// --- Siemens Structured Format ---
DATA_BLOCK "model_HS16_IW10"
{ S7_Optimized_Access := 'TRUE' }
VERSION : 0.1
NON_RETAIN
   VAR
      W_i : ARRAY[0..15, 0..39] OF REAL;
      W_f : ARRAY[0..15, 0..39] OF REAL;
      W_g : ARRAY[0..15, 0..39] OF REAL;
      W_o : ARRAY[0..15, 0..39] OF REAL;
      R_i : ARRAY[0..15, 0..15] OF REAL;
      R_f : ARRAY[0..15, 0..15] OF REAL;
      R_g : ARRAY[0..15, 0..15] OF REAL;
      R_o : ARRAY[0..15, 0..15] OF REAL;
      B_i : ARRAY[0..15] OF REAL;
      B_f : ARRAY[0..15] OF REAL;
      B_g : ARRAY[0..15] OF REAL;
      B_o : ARRAY[0..15] OF REAL;
      FC_W : ARRAY[0..39, 0..15] OF REAL;
      FC_B : ARRAY[0..39] OF REAL;
   END_VAR
BEGIN

      W_i[0,0] := 0.03254747;
      W_i[0,1] := 0.12385904;
      W_i[0,2] := 0.04015401;
      W_i[0,3] := -0.03803189;
      W_i[0,4] := 0.17593189;
      W_i[0,5] := 0.00417833;
      W_i[0,6] := -0.00157293;
      W_i[0,7] := 0.07286220;
      W_i[0,8] := 0.06175515;
      W_i[0,9] := -0.03080547;
      W_i[0,10] := 0.01361996;
      W_i[0,11] := -0.23670040;
      W_i[0,12] := 0.12512483;
      W_i[0,13] := -0.12038948;
      W_i[0,14] := 0.05234820;
      W_i[0,15] := 0.26305324;
      W_i[0,16] := -0.11475044;
      W_i[0,17] := 0.05957858;
      W_i[0,18] := -0.02271187;
      W_i[0,19] := -0.04982074;
      W_i[0,20] := 0.01270425;
      W_i[0,21] := 0.36205307;
      W_i[0,22] := -0.29144672;
      W_i[0,23] := 0.02366253;
      W_i[0,24] := -0.60242903;
      W_i[0,25] := -0.51985335;
      W_i[0,26] := 0.01890776;
      W_i[0,27] := -0.42442557;
      W_i[0,28] := 0.09802054;
      W_i[0,29] := -0.29197305;
      W_i[0,30] := 0.17564484;
      W_i[0,31] := -0.06584074;
      W_i[0,32] := 0.04272554;
      W_i[0,33] := 0.06813997;
      W_i[0,34] := 0.12439077;
      W_i[0,35] := -0.20625667;
      W_i[0,36] := 0.05875245;
      W_i[0,37] := -0.27000934;
      W_i[0,38] := 0.22123174;
      W_i[0,39] := 1.45426822;
      W_i[1,0] := 0.04402059;
      W_i[1,1] := 0.10076170;
      W_i[1,2] := -0.00997876;
      W_i[1,3] := 0.00796912;
      W_i[1,4] := -0.00383734;
      W_i[1,5] := -0.00800767;
      W_i[1,6] := 0.12291239;
      W_i[1,7] := 0.04417216;
      W_i[1,8] := -0.00160155;
      W_i[1,9] := -0.03973384;
      W_i[1,10] := -0.05576275;
      W_i[1,11] := 0.01415846;
      W_i[1,12] := -0.11022115;
      W_i[1,13] := 0.03613710;
      W_i[1,14] := -0.00464776;
      W_i[1,15] := -0.02071899;
      W_i[1,16] := 0.01651780;
      W_i[1,17] := -0.00011115;
      W_i[1,18] := 0.04986879;
      W_i[1,19] := -0.05042609;
      W_i[1,20] := 0.08610544;
      W_i[1,21] := 0.05673008;
      W_i[1,22] := -0.00434864;
      W_i[1,23] := 0.01197722;
      W_i[1,24] := -0.54585391;
      W_i[1,25] := -0.68996310;
      W_i[1,26] := 0.01104975;
      W_i[1,27] := 0.01825110;
      W_i[1,28] := 0.04478757;
      W_i[1,29] := -0.05586376;
      W_i[1,30] := 0.02979602;
      W_i[1,31] := 0.00707946;
      W_i[1,32] := 0.14649346;
      W_i[1,33] := 0.04832766;
      W_i[1,34] := -0.92027420;
      W_i[1,35] := -0.19189121;
      W_i[1,36] := 0.02485085;
      W_i[1,37] := -0.05241579;
      W_i[1,38] := 0.01553158;
      W_i[1,39] := -0.00394726;
      W_i[2,0] := 0.06704360;
      W_i[2,1] := -0.11752029;
      W_i[2,2] := 0.02326228;
      W_i[2,3] := -0.14317727;
      W_i[2,4] := -0.05582308;
      W_i[2,5] := 0.03605313;
      W_i[2,6] := 0.04952687;
      W_i[2,7] := -0.05419854;
      W_i[2,8] := -0.00077774;
      W_i[2,9] := 0.17699891;
      W_i[2,10] := 0.02469403;
      W_i[2,11] := 0.28494063;
      W_i[2,12] := -0.27127108;
      W_i[2,13] := -0.06837726;
      W_i[2,14] := 0.00509281;
      W_i[2,15] := 0.07467768;
      W_i[2,16] := 0.01470727;
      W_i[2,17] := 0.11394187;
      W_i[2,18] := -0.03895494;
      W_i[2,19] := 0.02999579;
      W_i[2,20] := 0.01967140;
      W_i[2,21] := 0.00220801;
      W_i[2,22] := -0.33803001;
      W_i[2,23] := 0.09799825;
      W_i[2,24] := -0.59557176;
      W_i[2,25] := -0.72284853;
      W_i[2,26] := 0.07928592;
      W_i[2,27] := -0.03053538;
      W_i[2,28] := -0.13099378;
      W_i[2,29] := -0.04490006;
      W_i[2,30] := 0.05262627;
      W_i[2,31] := -0.03356259;
      W_i[2,32] := 0.06378829;
      W_i[2,33] := -0.00362085;
      W_i[2,34] := -0.65794659;
      W_i[2,35] := 0.02030313;
      W_i[2,36] := 0.05807094;
      W_i[2,37] := -0.11176150;
      W_i[2,38] := 0.09806133;
      W_i[2,39] := -0.04513157;
      W_i[3,0] := -0.03288125;
      W_i[3,1] := 0.03644303;
      W_i[3,2] := -0.02111984;
      W_i[3,3] := -0.09554495;
      W_i[3,4] := 0.47103399;
      W_i[3,5] := -0.01821760;
      W_i[3,6] := -0.01296977;
      W_i[3,7] := 0.09772011;
      W_i[3,8] := 0.02375359;
      W_i[3,9] := 0.08029480;
      W_i[3,10] := 0.06341432;
      W_i[3,11] := -0.05777879;
      W_i[3,12] := 0.09200994;
      W_i[3,13] := -0.00543420;
      W_i[3,14] := -0.11079636;
      W_i[3,15] := 0.18567836;
      W_i[3,16] := -0.01795590;
      W_i[3,17] := -0.01424691;
      W_i[3,18] := 0.02418556;
      W_i[3,19] := -0.08783326;
      W_i[3,20] := 0.05560731;
      W_i[3,21] := 0.29868218;
      W_i[3,22] := -0.22202586;
      W_i[3,23] := -0.03734203;
      W_i[3,24] := 0.08825689;
      W_i[3,25] := 0.18388928;
      W_i[3,26] := 0.11525851;
      W_i[3,27] := -0.44497600;
      W_i[3,28] := 0.10198013;
      W_i[3,29] := -0.44026142;
      W_i[3,30] := -0.20704049;
      W_i[3,31] := 0.00454621;
      W_i[3,32] := -0.03864358;
      W_i[3,33] := -0.10321955;
      W_i[3,34] := 0.61782306;
      W_i[3,35] := -0.01621445;
      W_i[3,36] := 0.06078746;
      W_i[3,37] := 0.07829241;
      W_i[3,38] := 0.08872399;
      W_i[3,39] := 0.01815886;
      W_i[4,0] := -0.09336383;
      W_i[4,1] := 0.00870158;
      W_i[4,2] := -0.05045110;
      W_i[4,3] := 0.06854370;
      W_i[4,4] := 0.06657482;
      W_i[4,5] := -0.04358229;
      W_i[4,6] := 0.01173393;
      W_i[4,7] := 0.02832152;
      W_i[4,8] := -0.23808675;
      W_i[4,9] := 0.25903443;
      W_i[4,10] := -0.02959821;
      W_i[4,11] := -0.19702840;
      W_i[4,12] := -0.04782372;
      W_i[4,13] := 0.00693473;
      W_i[4,14] := 0.00193878;
      W_i[4,15] := 0.03396931;
      W_i[4,16] := -0.03933699;
      W_i[4,17] := -0.09345319;
      W_i[4,18] := 0.85718733;
      W_i[4,19] := -0.20839401;
      W_i[4,20] := -0.00447866;
      W_i[4,21] := -0.04350503;
      W_i[4,22] := 0.09176219;
      W_i[4,23] := 0.04992297;
      W_i[4,24] := -0.45042995;
      W_i[4,25] := 0.01641427;
      W_i[4,26] := -0.18378316;
      W_i[4,27] := 0.03955682;
      W_i[4,28] := -0.06913128;
      W_i[4,29] := 0.08025265;
      W_i[4,30] := -0.11622916;
      W_i[4,31] := 0.04558431;
      W_i[4,32] := 0.07176397;
      W_i[4,33] := -0.04032118;
      W_i[4,34] := 0.20981206;
      W_i[4,35] := -0.11253353;
      W_i[4,36] := -0.01868857;
      W_i[4,37] := -0.07242457;
      W_i[4,38] := -0.13242386;
      W_i[4,39] := -0.04244877;
      W_i[5,0] := 0.01391891;
      W_i[5,1] := -0.11018298;
      W_i[5,2] := -0.00893384;
      W_i[5,3] := -0.01407803;
      W_i[5,4] := 0.08575681;
      W_i[5,5] := 0.08241521;
      W_i[5,6] := -0.06153676;
      W_i[5,7] := 0.03060099;
      W_i[5,8] := -0.03490681;
      W_i[5,9] := 0.03142790;
      W_i[5,10] := -0.02459875;
      W_i[5,11] := 0.10959067;
      W_i[5,12] := -0.02965787;
      W_i[5,13] := 0.00184801;
      W_i[5,14] := 0.02055808;
      W_i[5,15] := -0.00937524;
      W_i[5,16] := -0.01257727;
      W_i[5,17] := 0.01791891;
      W_i[5,18] := -0.01156250;
      W_i[5,19] := -0.02731706;
      W_i[5,20] := 0.08900256;
      W_i[5,21] := 0.09895428;
      W_i[5,22] := 0.02720478;
      W_i[5,23] := 0.04369688;
      W_i[5,24] := -1.90607393;
      W_i[5,25] := -0.09418426;
      W_i[5,26] := -0.01059700;
      W_i[5,27] := -0.09780212;
      W_i[5,28] := 0.11255830;
      W_i[5,29] := 0.08197493;
      W_i[5,30] := -0.08072126;
      W_i[5,31] := 0.03083795;
      W_i[5,32] := 0.06895962;
      W_i[5,33] := 0.00149198;
      W_i[5,34] := 0.30098182;
      W_i[5,35] := 0.14424579;
      W_i[5,36] := -0.02817895;
      W_i[5,37] := -0.08498497;
      W_i[5,38] := 0.03758771;
      W_i[5,39] := 0.01095005;
      W_i[6,0] := 0.08324189;
      W_i[6,1] := -0.28836685;
      W_i[6,2] := -0.00092833;
      W_i[6,3] := -0.00874277;
      W_i[6,4] := 0.11969821;
      W_i[6,5] := -0.11207853;
      W_i[6,6] := -0.00877090;
      W_i[6,7] := -0.03745995;
      W_i[6,8] := 0.00287988;
      W_i[6,9] := 0.00178848;
      W_i[6,10] := 0.03823818;
      W_i[6,11] := 0.02621512;
      W_i[6,12] := -0.28842098;
      W_i[6,13] := -0.07084718;
      W_i[6,14] := 0.04070705;
      W_i[6,15] := -0.02042400;
      W_i[6,16] := -0.00164282;
      W_i[6,17] := 0.01065832;
      W_i[6,18] := 0.00655926;
      W_i[6,19] := 0.02358968;
      W_i[6,20] := 0.13037887;
      W_i[6,21] := 0.03868100;
      W_i[6,22] := -0.06235948;
      W_i[6,23] := 0.07983913;
      W_i[6,24] := -0.24280079;
      W_i[6,25] := -0.05732525;
      W_i[6,26] := 0.16517149;
      W_i[6,27] := -0.07414961;
      W_i[6,28] := 0.06032364;
      W_i[6,29] := 0.08282514;
      W_i[6,30] := -0.01358633;
      W_i[6,31] := 0.04311090;
      W_i[6,32] := 0.03472897;
      W_i[6,33] := -0.04253995;
      W_i[6,34] := 0.01447233;
      W_i[6,35] := 0.03594886;
      W_i[6,36] := -0.01385077;
      W_i[6,37] := 0.11164505;
      W_i[6,38] := 0.12532353;
      W_i[6,39] := -0.03726343;
      W_i[7,0] := 0.01927893;
      W_i[7,1] := 0.05625859;
      W_i[7,2] := 0.04672581;
      W_i[7,3] := -0.00316564;
      W_i[7,4] := 0.09401099;
      W_i[7,5] := -0.02755413;
      W_i[7,6] := -0.03952036;
      W_i[7,7] := 0.03364034;
      W_i[7,8] := 0.05500693;
      W_i[7,9] := 0.02471298;
      W_i[7,10] := 0.03820876;
      W_i[7,11] := -0.26921606;
      W_i[7,12] := -0.02231521;
      W_i[7,13] := -0.01752430;
      W_i[7,14] := 0.03934914;
      W_i[7,15] := 0.01282423;
      W_i[7,16] := -0.08716010;
      W_i[7,17] := -0.09125534;
      W_i[7,18] := 0.00613662;
      W_i[7,19] := 0.08651425;
      W_i[7,20] := -0.01288831;
      W_i[7,21] := 0.20176773;
      W_i[7,22] := -0.20166723;
      W_i[7,23] := 0.01241351;
      W_i[7,24] := -0.87556225;
      W_i[7,25] := -0.46218389;
      W_i[7,26] := 0.09773878;
      W_i[7,27] := -0.12810560;
      W_i[7,28] := 0.04194518;
      W_i[7,29] := -0.03563948;
      W_i[7,30] := 0.08049577;
      W_i[7,31] := 0.04509509;
      W_i[7,32] := -0.11332804;
      W_i[7,33] := 0.10539962;
      W_i[7,34] := 0.24167158;
      W_i[7,35] := 0.04508473;
      W_i[7,36] := 0.00324964;
      W_i[7,37] := 0.22550038;
      W_i[7,38] := 0.17509922;
      W_i[7,39] := -0.77876335;
      W_i[8,0] := -0.03076644;
      W_i[8,1] := 0.03958185;
      W_i[8,2] := 0.05958826;
      W_i[8,3] := 0.00143461;
      W_i[8,4] := -0.03551066;
      W_i[8,5] := 0.06705590;
      W_i[8,6] := -0.00545013;
      W_i[8,7] := -0.11520024;
      W_i[8,8] := -0.04941865;
      W_i[8,9] := 0.00970779;
      W_i[8,10] := -0.02700928;
      W_i[8,11] := 0.12616971;
      W_i[8,12] := -0.23012702;
      W_i[8,13] := -0.13218109;
      W_i[8,14] := 0.10565390;
      W_i[8,15] := 0.03265957;
      W_i[8,16] := 0.01893855;
      W_i[8,17] := 0.05783269;
      W_i[8,18] := 0.04541522;
      W_i[8,19] := -0.17565091;
      W_i[8,20] := -0.03008310;
      W_i[8,21] := 0.02609591;
      W_i[8,22] := -0.11792074;
      W_i[8,23] := -0.03097328;
      W_i[8,24] := -1.12349439;
      W_i[8,25] := -0.10578562;
      W_i[8,26] := 0.11967086;
      W_i[8,27] := -0.19309855;
      W_i[8,28] := -0.04314341;
      W_i[8,29] := -0.02280886;
      W_i[8,30] := 0.09419166;
      W_i[8,31] := -0.00168002;
      W_i[8,32] := 0.17011297;
      W_i[8,33] := 0.12776379;
      W_i[8,34] := 0.00792190;
      W_i[8,35] := 0.00793266;
      W_i[8,36] := 0.02933485;
      W_i[8,37] := -0.04765635;
      W_i[8,38] := -0.05385318;
      W_i[8,39] := 1.04576063;
      W_i[9,0] := 0.15918908;
      W_i[9,1] := 0.04106269;
      W_i[9,2] := 0.02940365;
      W_i[9,3] := -0.02633034;
      W_i[9,4] := 0.06646424;
      W_i[9,5] := -0.06870057;
      W_i[9,6] := 0.00617184;
      W_i[9,7] := 0.01493581;
      W_i[9,8] := 0.00472299;
      W_i[9,9] := -0.18171085;
      W_i[9,10] := -0.00863580;
      W_i[9,11] := 0.11203966;
      W_i[9,12] := 0.03235663;
      W_i[9,13] := -0.00635904;
      W_i[9,14] := -0.00805719;
      W_i[9,15] := 0.03256573;
      W_i[9,16] := -0.02982800;
      W_i[9,17] := 0.02432551;
      W_i[9,18] := -0.04791717;
      W_i[9,19] := -0.03479305;
      W_i[9,20] := 0.02419964;
      W_i[9,21] := -0.00806570;
      W_i[9,22] := 0.00884045;
      W_i[9,23] := 0.00822151;
      W_i[9,24] := -0.46266055;
      W_i[9,25] := -0.24154246;
      W_i[9,26] := 0.10637723;
      W_i[9,27] := 0.00555547;
      W_i[9,28] := 0.00231378;
      W_i[9,29] := 0.17306480;
      W_i[9,30] := -0.14428723;
      W_i[9,31] := -0.01611738;
      W_i[9,32] := -0.15273547;
      W_i[9,33] := -0.03995335;
      W_i[9,34] := -0.60233766;
      W_i[9,35] := -0.06071381;
      W_i[9,36] := 0.01153921;
      W_i[9,37] := 0.15725203;
      W_i[9,38] := 0.04887648;
      W_i[9,39] := 0.03194974;
      W_i[10,0] := 0.00000571;
      W_i[10,1] := 0.02921890;
      W_i[10,2] := 0.03921259;
      W_i[10,3] := -0.10342362;
      W_i[10,4] := 0.04451175;
      W_i[10,5] := -0.01788418;
      W_i[10,6] := 0.06014212;
      W_i[10,7] := -0.12761596;
      W_i[10,8] := 0.10969678;
      W_i[10,9] := 0.13464272;
      W_i[10,10] := -0.07629871;
      W_i[10,11] := -1.31473470;
      W_i[10,12] := 0.97041023;
      W_i[10,13] := -0.02917644;
      W_i[10,14] := 0.26857987;
      W_i[10,15] := 0.06801854;
      W_i[10,16] := -0.22419471;
      W_i[10,17] := 0.26248446;
      W_i[10,18] := -0.16949444;
      W_i[10,19] := -0.11971024;
      W_i[10,20] := -0.15914336;
      W_i[10,21] := 0.18180194;
      W_i[10,22] := -0.44877753;
      W_i[10,23] := 0.05718501;
      W_i[10,24] := 0.77401525;
      W_i[10,25] := 0.61128056;
      W_i[10,26] := 0.00735129;
      W_i[10,27] := -0.08243502;
      W_i[10,28] := -0.03729297;
      W_i[10,29] := 0.16128409;
      W_i[10,30] := -0.02351914;
      W_i[10,31] := 0.10431249;
      W_i[10,32] := 0.05746254;
      W_i[10,33] := 0.08887602;
      W_i[10,34] := -0.39106452;
      W_i[10,35] := 0.22569241;
      W_i[10,36] := -0.13208193;
      W_i[10,37] := -0.16115883;
      W_i[10,38] := 0.27080455;
      W_i[10,39] := 0.62801355;
      W_i[11,0] := -0.05849513;
      W_i[11,1] := -0.03062119;
      W_i[11,2] := -0.00411083;
      W_i[11,3] := 0.00799791;
      W_i[11,4] := 0.08333463;
      W_i[11,5] := 0.02937987;
      W_i[11,6] := 0.06844535;
      W_i[11,7] := -0.01198280;
      W_i[11,8] := 0.05660131;
      W_i[11,9] := -0.14609326;
      W_i[11,10] := -0.01666861;
      W_i[11,11] := -0.06908122;
      W_i[11,12] := 0.15483312;
      W_i[11,13] := -0.00687739;
      W_i[11,14] := 0.01971146;
      W_i[11,15] := 0.13305922;
      W_i[11,16] := -0.02189317;
      W_i[11,17] := 0.00985993;
      W_i[11,18] := -0.14880668;
      W_i[11,19] := 0.01909257;
      W_i[11,20] := 0.03714932;
      W_i[11,21] := -0.02673176;
      W_i[11,22] := -0.02788893;
      W_i[11,23] := 0.11408952;
      W_i[11,24] := -0.37118840;
      W_i[11,25] := -0.08985706;
      W_i[11,26] := -0.11023268;
      W_i[11,27] := 0.05117378;
      W_i[11,28] := 0.08547711;
      W_i[11,29] := 0.12702477;
      W_i[11,30] := 0.10544877;
      W_i[11,31] := -0.00480978;
      W_i[11,32] := 0.16144946;
      W_i[11,33] := 0.05210381;
      W_i[11,34] := -0.00085451;
      W_i[11,35] := -0.00874526;
      W_i[11,36] := -0.06161120;
      W_i[11,37] := -0.36774832;
      W_i[11,38] := 0.04212995;
      W_i[11,39] := 0.03037546;
      W_i[12,0] := 0.00629061;
      W_i[12,1] := -0.06136212;
      W_i[12,2] := -0.00718669;
      W_i[12,3] := -0.10042179;
      W_i[12,4] := 0.06293897;
      W_i[12,5] := -0.03143417;
      W_i[12,6] := -0.03538829;
      W_i[12,7] := 0.07763195;
      W_i[12,8] := -0.01023159;
      W_i[12,9] := -0.11412965;
      W_i[12,10] := -0.01354402;
      W_i[12,11] := -0.02311977;
      W_i[12,12] := 0.02796080;
      W_i[12,13] := 0.07165248;
      W_i[12,14] := -0.03632027;
      W_i[12,15] := 0.03878558;
      W_i[12,16] := -0.07312500;
      W_i[12,17] := 0.01845204;
      W_i[12,18] := -0.08527449;
      W_i[12,19] := -0.00854577;
      W_i[12,20] := 0.00351815;
      W_i[12,21] := -0.16628480;
      W_i[12,22] := 0.06705266;
      W_i[12,23] := 0.14307018;
      W_i[12,24] := -0.53957397;
      W_i[12,25] := -0.87219816;
      W_i[12,26] := -0.06440469;
      W_i[12,27] := 0.07379381;
      W_i[12,28] := 0.07828815;
      W_i[12,29] := 0.38822088;
      W_i[12,30] := 0.11594980;
      W_i[12,31] := 0.05581488;
      W_i[12,32] := 0.30664018;
      W_i[12,33] := 0.12759578;
      W_i[12,34] := -0.14797799;
      W_i[12,35] := 0.14329346;
      W_i[12,36] := 0.22981535;
      W_i[12,37] := 0.00895516;
      W_i[12,38] := 0.20012984;
      W_i[12,39] := 0.09707437;
      W_i[13,0] := 0.07871004;
      W_i[13,1] := 0.06409820;
      W_i[13,2] := -0.00181766;
      W_i[13,3] := 0.05780525;
      W_i[13,4] := 0.21016718;
      W_i[13,5] := 0.05360549;
      W_i[13,6] := -0.08758270;
      W_i[13,7] := -0.33428112;
      W_i[13,8] := -0.09135646;
      W_i[13,9] := 0.11706311;
      W_i[13,10] := -0.05231260;
      W_i[13,11] := -0.03317479;
      W_i[13,12] := -0.40338296;
      W_i[13,13] := -0.00985299;
      W_i[13,14] := 0.02202887;
      W_i[13,15] := 0.13037799;
      W_i[13,16] := 0.04808246;
      W_i[13,17] := 0.04501719;
      W_i[13,18] := -0.01153503;
      W_i[13,19] := 0.03141625;
      W_i[13,20] := 0.02999944;
      W_i[13,21] := 0.01402024;
      W_i[13,22] := 0.06788336;
      W_i[13,23] := -0.09942459;
      W_i[13,24] := 0.31843993;
      W_i[13,25] := 0.10697926;
      W_i[13,26] := -0.06989229;
      W_i[13,27] := 0.10588147;
      W_i[13,28] := 0.06872193;
      W_i[13,29] := -0.15371445;
      W_i[13,30] := 0.06626805;
      W_i[13,31] := -0.05594840;
      W_i[13,32] := -0.09573574;
      W_i[13,33] := 0.05669653;
      W_i[13,34] := 0.06202357;
      W_i[13,35] := -0.13674185;
      W_i[13,36] := 0.06451428;
      W_i[13,37] := 0.12041676;
      W_i[13,38] := -0.16850901;
      W_i[13,39] := 0.97759265;
      W_i[14,0] := 0.00773311;
      W_i[14,1] := -0.06673568;
      W_i[14,2] := -0.03463669;
      W_i[14,3] := -0.07830913;
      W_i[14,4] := 0.22799005;
      W_i[14,5] := -0.23448689;
      W_i[14,6] := 0.19569355;
      W_i[14,7] := 0.13153341;
      W_i[14,8] := -0.12420856;
      W_i[14,9] := 0.28603974;
      W_i[14,10] := -0.09231006;
      W_i[14,11] := -0.25477913;
      W_i[14,12] := 0.14903630;
      W_i[14,13] := -0.29128024;
      W_i[14,14] := 0.10725706;
      W_i[14,15] := 0.13540378;
      W_i[14,16] := -0.09035023;
      W_i[14,17] := -0.01749873;
      W_i[14,18] := -0.47894967;
      W_i[14,19] := -0.06870104;
      W_i[14,20] := -0.17096391;
      W_i[14,21] := -0.05212005;
      W_i[14,22] := -0.16184741;
      W_i[14,23] := -0.21394062;
      W_i[14,24] := -0.75706887;
      W_i[14,25] := -0.70485926;
      W_i[14,26] := -0.33521020;
      W_i[14,27] := 0.03507431;
      W_i[14,28] := -0.12678961;
      W_i[14,29] := 0.16709636;
      W_i[14,30] := -0.05052740;
      W_i[14,31] := -0.11800393;
      W_i[14,32] := -0.09575160;
      W_i[14,33] := -0.01452094;
      W_i[14,34] := 0.00625472;
      W_i[14,35] := -0.12877558;
      W_i[14,36] := -0.06069501;
      W_i[14,37] := -0.22877042;
      W_i[14,38] := 0.17231728;
      W_i[14,39] := 1.04831111;
      W_i[15,0] := 0.04376059;
      W_i[15,1] := -0.02296846;
      W_i[15,2] := 0.01713722;
      W_i[15,3] := 0.17107451;
      W_i[15,4] := 0.17369278;
      W_i[15,5] := -0.01825109;
      W_i[15,6] := -0.02258963;
      W_i[15,7] := 0.02190229;
      W_i[15,8] := -0.03702974;
      W_i[15,9] := -0.03196403;
      W_i[15,10] := 0.08264420;
      W_i[15,11] := 0.05920084;
      W_i[15,12] := -0.42805931;
      W_i[15,13] := -0.17172982;
      W_i[15,14] := 0.02115602;
      W_i[15,15] := -0.00198027;
      W_i[15,16] := 0.02912534;
      W_i[15,17] := -0.07075519;
      W_i[15,18] := -0.11744455;
      W_i[15,19] := 0.30688557;
      W_i[15,20] := 0.04301663;
      W_i[15,21] := 0.21635388;
      W_i[15,22] := -0.08966552;
      W_i[15,23] := 0.07217173;
      W_i[15,24] := -0.53244919;
      W_i[15,25] := -0.17169446;
      W_i[15,26] := -0.00556448;
      W_i[15,27] := -0.16294074;
      W_i[15,28] := 0.03264420;
      W_i[15,29] := 0.01573053;
      W_i[15,30] := -0.03329111;
      W_i[15,31] := -0.01247096;
      W_i[15,32] := 0.21000683;
      W_i[15,33] := 0.15043637;
      W_i[15,34] := -0.16979790;
      W_i[15,35] := 0.00504174;
      W_i[15,36] := 0.00267995;
      W_i[15,37] := -0.06215737;
      W_i[15,38] := 0.21481486;
      W_i[15,39] := 0.07231134;
      W_f[0,0] := -0.02091779;
      W_f[0,1] := -0.01810063;
      W_f[0,2] := 0.21008702;
      W_f[0,3] := 0.09207959;
      W_f[0,4] := -0.10695104;
      W_f[0,5] := -0.03611851;
      W_f[0,6] := 0.03397696;
      W_f[0,7] := 0.16544856;
      W_f[0,8] := -0.05997881;
      W_f[0,9] := -0.00453302;
      W_f[0,10] := 0.03307042;
      W_f[0,11] := 0.14202486;
      W_f[0,12] := 0.08012222;
      W_f[0,13] := -0.01528266;
      W_f[0,14] := -0.15201145;
      W_f[0,15] := -0.15718380;
      W_f[0,16] := -0.08413183;
      W_f[0,17] := 0.20222495;
      W_f[0,18] := -0.01353853;
      W_f[0,19] := 0.02782044;
      W_f[0,20] := -0.04748038;
      W_f[0,21] := 0.18304287;
      W_f[0,22] := 0.31257400;
      W_f[0,23] := -0.06208337;
      W_f[0,24] := 1.60133708;
      W_f[0,25] := 1.51956844;
      W_f[0,26] := 0.00266673;
      W_f[0,27] := 0.12180892;
      W_f[0,28] := 0.04435247;
      W_f[0,29] := 0.03200248;
      W_f[0,30] := 0.38338348;
      W_f[0,31] := 0.04435838;
      W_f[0,32] := 0.30680922;
      W_f[0,33] := 0.13231254;
      W_f[0,34] := 1.35719514;
      W_f[0,35] := 0.36870065;
      W_f[0,36] := 0.08067872;
      W_f[0,37] := 0.21299456;
      W_f[0,38] := -0.02734181;
      W_f[0,39] := 0.07611577;
      W_f[1,0] := -0.38817102;
      W_f[1,1] := 0.02779610;
      W_f[1,2] := -0.26510856;
      W_f[1,3] := -0.07072625;
      W_f[1,4] := 0.11966246;
      W_f[1,5] := 0.12000409;
      W_f[1,6] := -0.50846916;
      W_f[1,7] := -0.13361093;
      W_f[1,8] := -0.13777961;
      W_f[1,9] := -0.08736181;
      W_f[1,10] := 0.31134772;
      W_f[1,11] := 0.08504082;
      W_f[1,12] := 0.21148330;
      W_f[1,13] := -0.13549544;
      W_f[1,14] := -0.12279948;
      W_f[1,15] := 0.05185516;
      W_f[1,16] := -0.14745373;
      W_f[1,17] := 0.05817819;
      W_f[1,18] := 1.08165765;
      W_f[1,19] := 0.18381153;
      W_f[1,20] := 0.28742057;
      W_f[1,21] := -0.27315989;
      W_f[1,22] := 0.08855448;
      W_f[1,23] := -0.09573217;
      W_f[1,24] := -0.36683315;
      W_f[1,25] := -0.69911557;
      W_f[1,26] := 0.07979747;
      W_f[1,27] := -0.17541142;
      W_f[1,28] := -0.24551585;
      W_f[1,29] := 0.14984873;
      W_f[1,30] := 0.02324941;
      W_f[1,31] := 0.07932284;
      W_f[1,32] := -0.12442444;
      W_f[1,33] := 0.02366536;
      W_f[1,34] := 0.13745289;
      W_f[1,35] := 0.46306115;
      W_f[1,36] := -0.22673251;
      W_f[1,37] := 0.07258049;
      W_f[1,38] := 0.42296681;
      W_f[1,39] := 0.14921528;
      W_f[2,0] := -0.01982149;
      W_f[2,1] := 0.03324119;
      W_f[2,2] := -0.04425151;
      W_f[2,3] := 0.08356856;
      W_f[2,4] := -0.00266197;
      W_f[2,5] := -0.01017811;
      W_f[2,6] := -0.03237398;
      W_f[2,7] := -0.00609645;
      W_f[2,8] := -0.04705935;
      W_f[2,9] := 0.03853706;
      W_f[2,10] := 0.03140420;
      W_f[2,11] := -0.12043314;
      W_f[2,12] := 0.26915759;
      W_f[2,13] := 0.04188414;
      W_f[2,14] := 0.10631428;
      W_f[2,15] := 0.05646345;
      W_f[2,16] := 0.16197611;
      W_f[2,17] := 0.21402863;
      W_f[2,18] := -0.09279267;
      W_f[2,19] := -0.00577110;
      W_f[2,20] := -0.03028176;
      W_f[2,21] := -0.05153098;
      W_f[2,22] := -0.11017115;
      W_f[2,23] := -0.01419843;
      W_f[2,24] := -0.63084757;
      W_f[2,25] := -0.41158974;
      W_f[2,26] := -0.14941035;
      W_f[2,27] := 0.04505387;
      W_f[2,28] := 0.09163468;
      W_f[2,29] := 0.20423372;
      W_f[2,30] := -0.05021087;
      W_f[2,31] := -0.05815214;
      W_f[2,32] := -0.04207016;
      W_f[2,33] := 0.21736744;
      W_f[2,34] := 0.64307344;
      W_f[2,35] := -0.19552369;
      W_f[2,36] := -0.05630085;
      W_f[2,37] := 0.00531330;
      W_f[2,38] := -0.12282822;
      W_f[2,39] := 0.54551679;
      W_f[3,0] := -0.00758014;
      W_f[3,1] := 0.00559481;
      W_f[3,2] := 0.04034248;
      W_f[3,3] := 0.02266315;
      W_f[3,4] := -0.09543922;
      W_f[3,5] := 0.03211372;
      W_f[3,6] := 0.07329436;
      W_f[3,7] := -0.04057672;
      W_f[3,8] := -0.09598581;
      W_f[3,9] := -0.00159119;
      W_f[3,10] := 0.00039486;
      W_f[3,11] := -0.00788106;
      W_f[3,12] := -0.06210583;
      W_f[3,13] := -0.01413072;
      W_f[3,14] := -0.24013861;
      W_f[3,15] := -0.07759018;
      W_f[3,16] := 0.04360460;
      W_f[3,17] := -0.20987833;
      W_f[3,18] := 0.14860362;
      W_f[3,19] := -0.02982033;
      W_f[3,20] := -0.08417022;
      W_f[3,21] := 0.08484244;
      W_f[3,22] := 0.33418563;
      W_f[3,23] := -0.01567571;
      W_f[3,24] := 1.09344435;
      W_f[3,25] := 0.97723728;
      W_f[3,26] := -0.13622019;
      W_f[3,27] := -0.09956130;
      W_f[3,28] := 0.00698416;
      W_f[3,29] := 0.00054130;
      W_f[3,30] := 0.26053473;
      W_f[3,31] := -0.09947061;
      W_f[3,32] := 0.26287073;
      W_f[3,33] := 0.00611334;
      W_f[3,34] := 1.38905013;
      W_f[3,35] := -0.14349753;
      W_f[3,36] := -0.00342261;
      W_f[3,37] := -0.06542191;
      W_f[3,38] := 0.10482345;
      W_f[3,39] := 0.11385954;
      W_f[4,0] := 0.28678942;
      W_f[4,1] := -0.14550023;
      W_f[4,2] := 0.20301139;
      W_f[4,3] := -0.15284956;
      W_f[4,4] := -0.11934043;
      W_f[4,5] := -0.06261637;
      W_f[4,6] := -0.09047025;
      W_f[4,7] := -0.02217131;
      W_f[4,8] := 0.32893139;
      W_f[4,9] := -0.50192183;
      W_f[4,10] := -0.02496753;
      W_f[4,11] := -0.02753776;
      W_f[4,12] := -0.31547716;
      W_f[4,13] := -0.04408565;
      W_f[4,14] := 0.05384916;
      W_f[4,15] := -0.32536885;
      W_f[4,16] := -0.01380023;
      W_f[4,17] := -0.12124701;
      W_f[4,18] := 0.62146658;
      W_f[4,19] := 0.01393374;
      W_f[4,20] := 0.04359875;
      W_f[4,21] := 0.16302615;
      W_f[4,22] := -0.21024738;
      W_f[4,23] := -0.12911762;
      W_f[4,24] := -0.08685920;
      W_f[4,25] := -0.03674764;
      W_f[4,26] := 0.30872664;
      W_f[4,27] := 0.03806484;
      W_f[4,28] := 0.01020021;
      W_f[4,29] := -0.15197505;
      W_f[4,30] := 0.05839425;
      W_f[4,31] := -0.01564794;
      W_f[4,32] := -0.18343291;
      W_f[4,33] := 0.02443381;
      W_f[4,34] := 0.21402271;
      W_f[4,35] := 0.19360679;
      W_f[4,36] := 0.09160208;
      W_f[4,37] := 0.06046678;
      W_f[4,38] := -0.08968955;
      W_f[4,39] := -0.03439303;
      W_f[5,0] := -0.39957133;
      W_f[5,1] := -0.46507514;
      W_f[5,2] := -0.26463589;
      W_f[5,3] := -0.08991144;
      W_f[5,4] := -0.16602752;
      W_f[5,5] := 0.36502278;
      W_f[5,6] := -0.03514609;
      W_f[5,7] := -0.06387420;
      W_f[5,8] := 0.12637840;
      W_f[5,9] := 0.19450709;
      W_f[5,10] := -0.07852599;
      W_f[5,11] := -0.24370454;
      W_f[5,12] := -0.06879438;
      W_f[5,13] := 0.26811865;
      W_f[5,14] := 0.01808503;
      W_f[5,15] := -0.10070925;
      W_f[5,16] := 0.31043285;
      W_f[5,17] := -0.03764273;
      W_f[5,18] := -0.05466426;
      W_f[5,19] := -0.10286047;
      W_f[5,20] := -0.18913145;
      W_f[5,21] := -0.06289500;
      W_f[5,22] := 0.26261428;
      W_f[5,23] := 0.11659861;
      W_f[5,24] := 2.13931274;
      W_f[5,25] := 2.36269403;
      W_f[5,26] := -0.41290748;
      W_f[5,27] := 0.08711372;
      W_f[5,28] := -0.06960621;
      W_f[5,29] := -0.10882857;
      W_f[5,30] := 0.02405319;
      W_f[5,31] := -0.02791615;
      W_f[5,32] := -0.03174478;
      W_f[5,33] := -0.22598031;
      W_f[5,34] := 0.02213258;
      W_f[5,35] := 0.06206211;
      W_f[5,36] := -0.22062500;
      W_f[5,37] := 0.20298730;
      W_f[5,38] := 0.03730853;
      W_f[5,39] := -0.16448267;
      W_f[6,0] := 0.09157378;
      W_f[6,1] := -0.10600298;
      W_f[6,2] := 0.01516851;
      W_f[6,3] := -0.09814398;
      W_f[6,4] := -0.02060772;
      W_f[6,5] := -0.11663528;
      W_f[6,6] := 0.17605469;
      W_f[6,7] := 0.14043835;
      W_f[6,8] := -0.06626645;
      W_f[6,9] := 0.03254180;
      W_f[6,10] := -0.03667779;
      W_f[6,11] := 0.03295979;
      W_f[6,12] := 0.13456115;
      W_f[6,13] := 0.17527823;
      W_f[6,14] := 0.06438499;
      W_f[6,15] := -0.12721057;
      W_f[6,16] := -0.28780875;
      W_f[6,17] := 0.11614764;
      W_f[6,18] := -0.23114346;
      W_f[6,19] := -0.07521003;
      W_f[6,20] := -0.14160164;
      W_f[6,21] := 0.12687035;
      W_f[6,22] := 0.38557813;
      W_f[6,23] := -0.12900937;
      W_f[6,24] := 1.14550745;
      W_f[6,25] := 1.20651269;
      W_f[6,26] := 0.01718643;
      W_f[6,27] := -0.20140134;
      W_f[6,28] := -0.03907681;
      W_f[6,29] := -1.03183591;
      W_f[6,30] := 0.13298695;
      W_f[6,31] := -0.05304611;
      W_f[6,32] := 0.27542382;
      W_f[6,33] := 0.48400101;
      W_f[6,34] := 0.87303483;
      W_f[6,35] := -0.27916309;
      W_f[6,36] := 0.09285419;
      W_f[6,37] := -0.00086587;
      W_f[6,38] := 0.21403548;
      W_f[6,39] := 0.01036415;
      W_f[7,0] := -0.00185265;
      W_f[7,1] := 0.07858364;
      W_f[7,2] := 0.00610039;
      W_f[7,3] := 0.06575946;
      W_f[7,4] := -0.08100830;
      W_f[7,5] := 0.00321988;
      W_f[7,6] := 0.07597861;
      W_f[7,7] := -0.12638623;
      W_f[7,8] := 0.14672390;
      W_f[7,9] := 0.04145058;
      W_f[7,10] := 0.03552409;
      W_f[7,11] := -0.42004111;
      W_f[7,12] := 0.25357988;
      W_f[7,13] := -0.08330481;
      W_f[7,14] := -0.08974353;
      W_f[7,15] := -0.10517624;
      W_f[7,16] := -0.38224444;
      W_f[7,17] := -0.45799860;
      W_f[7,18] := -0.06309059;
      W_f[7,19] := -0.30799860;
      W_f[7,20] := -0.08522949;
      W_f[7,21] := -0.06581733;
      W_f[7,22] := 0.25805131;
      W_f[7,23] := 0.02311642;
      W_f[7,24] := 0.90950686;
      W_f[7,25] := 1.18889558;
      W_f[7,26] := -0.11546607;
      W_f[7,27] := -0.10872247;
      W_f[7,28] := -0.08876549;
      W_f[7,29] := 0.00109644;
      W_f[7,30] := 0.23372188;
      W_f[7,31] := -0.13769329;
      W_f[7,32] := 0.16597158;
      W_f[7,33] := 0.04170239;
      W_f[7,34] := 1.31133747;
      W_f[7,35] := -0.11888772;
      W_f[7,36] := 0.04907094;
      W_f[7,37] := 0.14026117;
      W_f[7,38] := 0.12559824;
      W_f[7,39] := -1.27418923;
      W_f[8,0] := 0.12555996;
      W_f[8,1] := -0.10315757;
      W_f[8,2] := 0.03551091;
      W_f[8,3] := -0.03898631;
      W_f[8,4] := -0.13206761;
      W_f[8,5] := 0.07454634;
      W_f[8,6] := 0.10206546;
      W_f[8,7] := 0.01262685;
      W_f[8,8] := -0.00534601;
      W_f[8,9] := -0.00536494;
      W_f[8,10] := -0.04092396;
      W_f[8,11] := -0.38692373;
      W_f[8,12] := 0.03422466;
      W_f[8,13] := 0.02580789;
      W_f[8,14] := 0.26898870;
      W_f[8,15] := -0.24944888;
      W_f[8,16] := -0.02722716;
      W_f[8,17] := -0.10108043;
      W_f[8,18] := 0.54244351;
      W_f[8,19] := -0.23120664;
      W_f[8,20] := -0.04103015;
      W_f[8,21] := -0.16740812;
      W_f[8,22] := 0.13893805;
      W_f[8,23] := -0.04656294;
      W_f[8,24] := 0.53174204;
      W_f[8,25] := 0.74309415;
      W_f[8,26] := -0.00084738;
      W_f[8,27] := -0.04600925;
      W_f[8,28] := -0.15880004;
      W_f[8,29] := 0.08535929;
      W_f[8,30] := 0.10221286;
      W_f[8,31] := -0.03335671;
      W_f[8,32] := 0.03138823;
      W_f[8,33] := -0.02403146;
      W_f[8,34] := 0.83305961;
      W_f[8,35] := -0.07033388;
      W_f[8,36] := -0.17499864;
      W_f[8,37] := 0.09229370;
      W_f[8,38] := -0.17668678;
      W_f[8,39] := 0.14198503;
      W_f[9,0] := -0.08198071;
      W_f[9,1] := 0.03835172;
      W_f[9,2] := 1.02026522;
      W_f[9,3] := -0.15293953;
      W_f[9,4] := -0.16179894;
      W_f[9,5] := 0.03072036;
      W_f[9,6] := -0.09759208;
      W_f[9,7] := -0.07946933;
      W_f[9,8] := -0.65491873;
      W_f[9,9] := 0.24554865;
      W_f[9,10] := -0.00084776;
      W_f[9,11] := -0.02393647;
      W_f[9,12] := -0.11035760;
      W_f[9,13] := 0.05757844;
      W_f[9,14] := 0.00252463;
      W_f[9,15] := -0.04278835;
      W_f[9,16] := -0.01363701;
      W_f[9,17] := 0.03181182;
      W_f[9,18] := 0.29542166;
      W_f[9,19] := 0.18680713;
      W_f[9,20] := -0.14596237;
      W_f[9,21] := 0.04626612;
      W_f[9,22] := -0.49596560;
      W_f[9,23] := -0.29882804;
      W_f[9,24] := -0.05025842;
      W_f[9,25] := -0.24922217;
      W_f[9,26] := 0.22770426;
      W_f[9,27] := -0.07712200;
      W_f[9,28] := -0.16018625;
      W_f[9,29] := -0.36028501;
      W_f[9,30] := -0.15894593;
      W_f[9,31] := 0.07634185;
      W_f[9,32] := -0.14248089;
      W_f[9,33] := 0.47243714;
      W_f[9,34] := 0.37227076;
      W_f[9,35] := 0.08862774;
      W_f[9,36] := 0.18020450;
      W_f[9,37] := -0.46372715;
      W_f[9,38] := 0.10143350;
      W_f[9,39] := 0.03257460;
      W_f[10,0] := 0.01476683;
      W_f[10,1] := 0.08915940;
      W_f[10,2] := 0.09493639;
      W_f[10,3] := 0.00921640;
      W_f[10,4] := -0.40101719;
      W_f[10,5] := -0.09464957;
      W_f[10,6] := -0.04691195;
      W_f[10,7] := -0.02866868;
      W_f[10,8] := -0.04315028;
      W_f[10,9] := -0.17093825;
      W_f[10,10] := -0.00073274;
      W_f[10,11] := -0.27505547;
      W_f[10,12] := 0.33605671;
      W_f[10,13] := -0.22034417;
      W_f[10,14] := 0.24165145;
      W_f[10,15] := -0.23521844;
      W_f[10,16] := -0.00154005;
      W_f[10,17] := -0.00158511;
      W_f[10,18] := 0.11912328;
      W_f[10,19] := -0.02448388;
      W_f[10,20] := -0.23859039;
      W_f[10,21] := -0.05945824;
      W_f[10,22] := 0.01714438;
      W_f[10,23] := -0.18285508;
      W_f[10,24] := 1.57859039;
      W_f[10,25] := 1.89422643;
      W_f[10,26] := 0.09559432;
      W_f[10,27] := -0.27382705;
      W_f[10,28] := -0.28146487;
      W_f[10,29] := 0.04344108;
      W_f[10,30] := 0.08430442;
      W_f[10,31] := 0.13571435;
      W_f[10,32] := 0.03089454;
      W_f[10,33] := 0.19871859;
      W_f[10,34] := 0.12124728;
      W_f[10,35] := 0.13877974;
      W_f[10,36] := 0.26381519;
      W_f[10,37] := 0.00209056;
      W_f[10,38] := -0.08942132;
      W_f[10,39] := -0.44943866;
      W_f[11,0] := 0.04211291;
      W_f[11,1] := -0.02505053;
      W_f[11,2] := 0.08745301;
      W_f[11,3] := -0.04265523;
      W_f[11,4] := -0.21276116;
      W_f[11,5] := 0.01322894;
      W_f[11,6] := 0.10620508;
      W_f[11,7] := 0.01512342;
      W_f[11,8] := -0.07057641;
      W_f[11,9] := 0.12398467;
      W_f[11,10] := -0.14091872;
      W_f[11,11] := -0.07267960;
      W_f[11,12] := 0.00417219;
      W_f[11,13] := -0.01783882;
      W_f[11,14] := 0.01799064;
      W_f[11,15] := -0.05493079;
      W_f[11,16] := -0.05114271;
      W_f[11,17] := -0.03128599;
      W_f[11,18] := 0.03801877;
      W_f[11,19] := -0.01814952;
      W_f[11,20] := -0.09758195;
      W_f[11,21] := -0.04573784;
      W_f[11,22] := -0.03167154;
      W_f[11,23] := -0.08901857;
      W_f[11,24] := -0.22173922;
      W_f[11,25] := 0.39944053;
      W_f[11,26] := 0.05129110;
      W_f[11,27] := 0.05733421;
      W_f[11,28] := -0.12204757;
      W_f[11,29] := 0.25301519;
      W_f[11,30] := -0.01943143;
      W_f[11,31] := 0.06523979;
      W_f[11,32] := -0.19657055;
      W_f[11,33] := 0.01042900;
      W_f[11,34] := 0.19335911;
      W_f[11,35] := -0.02032585;
      W_f[11,36] := -0.05446678;
      W_f[11,37] := 0.10930583;
      W_f[11,38] := -0.05791799;
      W_f[11,39] := 0.32721651;
      W_f[12,0] := 0.05839740;
      W_f[12,1] := 0.06337267;
      W_f[12,2] := 0.05269343;
      W_f[12,3] := -0.02425898;
      W_f[12,4] := 0.07333850;
      W_f[12,5] := 0.01520942;
      W_f[12,6] := 0.03044897;
      W_f[12,7] := 0.11511354;
      W_f[12,8] := 0.03681342;
      W_f[12,9] := -0.01680350;
      W_f[12,10] := 0.04408923;
      W_f[12,11] := 0.08383411;
      W_f[12,12] := -0.01220268;
      W_f[12,13] := 0.05396410;
      W_f[12,14] := -0.07032214;
      W_f[12,15] := -0.00997462;
      W_f[12,16] := -0.06021495;
      W_f[12,17] := -0.01422043;
      W_f[12,18] := -0.00584967;
      W_f[12,19] := 0.05498984;
      W_f[12,20] := -0.09216670;
      W_f[12,21] := 0.10788208;
      W_f[12,22] := 0.09067565;
      W_f[12,23] := -0.09486815;
      W_f[12,24] := -0.87601417;
      W_f[12,25] := 0.54372799;
      W_f[12,26] := 0.04737720;
      W_f[12,27] := -0.10040826;
      W_f[12,28] := 0.07258554;
      W_f[12,29] := 0.07306878;
      W_f[12,30] := -0.14698188;
      W_f[12,31] := 0.01059632;
      W_f[12,32] := 0.01764544;
      W_f[12,33] := -0.04630747;
      W_f[12,34] := 0.04829778;
      W_f[12,35] := -0.00637231;
      W_f[12,36] := 0.34302515;
      W_f[12,37] := 0.12217984;
      W_f[12,38] := 0.04078831;
      W_f[12,39] := 0.02011232;
      W_f[13,0] := 0.15987755;
      W_f[13,1] := 0.08477814;
      W_f[13,2] := -0.11990058;
      W_f[13,3] := -0.21518369;
      W_f[13,4] := 0.04422749;
      W_f[13,5] := 0.16439709;
      W_f[13,6] := -0.01991516;
      W_f[13,7] := 0.01602156;
      W_f[13,8] := -0.13440605;
      W_f[13,9] := 0.04321520;
      W_f[13,10] := 0.12583691;
      W_f[13,11] := 0.03486055;
      W_f[13,12] := 0.18403338;
      W_f[13,13] := 0.05531228;
      W_f[13,14] := -0.05205994;
      W_f[13,15] := -0.14179915;
      W_f[13,16] := 0.21455689;
      W_f[13,17] := -0.03670088;
      W_f[13,18] := 0.05554622;
      W_f[13,19] := -0.07012140;
      W_f[13,20] := 0.05645064;
      W_f[13,21] := 0.04904451;
      W_f[13,22] := 0.12274069;
      W_f[13,23] := -0.13912246;
      W_f[13,24] := 1.28141677;
      W_f[13,25] := 1.15295243;
      W_f[13,26] := 0.02036783;
      W_f[13,27] := 0.00000646;
      W_f[13,28] := 0.05594068;
      W_f[13,29] := 0.11384209;
      W_f[13,30] := 0.23915862;
      W_f[13,31] := 0.04423625;
      W_f[13,32] := 0.37905067;
      W_f[13,33] := 0.01350218;
      W_f[13,34] := 0.90777701;
      W_f[13,35] := -0.01705103;
      W_f[13,36] := 0.08728553;
      W_f[13,37] := 0.13768719;
      W_f[13,38] := 0.05409899;
      W_f[13,39] := 0.58763230;
      W_f[14,0] := -0.18308778;
      W_f[14,1] := 0.00258858;
      W_f[14,2] := -0.05409549;
      W_f[14,3] := 0.42653167;
      W_f[14,4] := -0.16614716;
      W_f[14,5] := -0.06032855;
      W_f[14,6] := 0.09126755;
      W_f[14,7] := -0.16223437;
      W_f[14,8] := -0.04155440;
      W_f[14,9] := -0.03031821;
      W_f[14,10] := -0.07388397;
      W_f[14,11] := -0.16659716;
      W_f[14,12] := 0.12239914;
      W_f[14,13] := -0.13348925;
      W_f[14,14] := -0.06961614;
      W_f[14,15] := -0.04957403;
      W_f[14,16] := 0.02988490;
      W_f[14,17] := -0.13393891;
      W_f[14,18] := -0.04285705;
      W_f[14,19] := -0.08629614;
      W_f[14,20] := -0.15329672;
      W_f[14,21] := 0.04812383;
      W_f[14,22] := -0.03088393;
      W_f[14,23] := -0.04624541;
      W_f[14,24] := -0.07781153;
      W_f[14,25] := -0.83196443;
      W_f[14,26] := 0.10154009;
      W_f[14,27] := 0.04807844;
      W_f[14,28] := 0.08697836;
      W_f[14,29] := -0.30993941;
      W_f[14,30] := 0.02526759;
      W_f[14,31] := 0.06875665;
      W_f[14,32] := 0.05270454;
      W_f[14,33] := 0.08052166;
      W_f[14,34] := 0.07316659;
      W_f[14,35] := -0.22593051;
      W_f[14,36] := -0.03604140;
      W_f[14,37] := -0.11075277;
      W_f[14,38] := 0.14222871;
      W_f[14,39] := 0.11912529;
      W_f[15,0] := 0.06860624;
      W_f[15,1] := 0.21167134;
      W_f[15,2] := -0.10700771;
      W_f[15,3] := -0.17963767;
      W_f[15,4] := 0.06190439;
      W_f[15,5] := 0.11186377;
      W_f[15,6] := 0.21238039;
      W_f[15,7] := 0.04805397;
      W_f[15,8] := 0.02383129;
      W_f[15,9] := -0.08112741;
      W_f[15,10] := -0.00035556;
      W_f[15,11] := -0.00759834;
      W_f[15,12] := 0.04278949;
      W_f[15,13] := -0.01575772;
      W_f[15,14] := -0.06780741;
      W_f[15,15] := 0.07988951;
      W_f[15,16] := 0.35835415;
      W_f[15,17] := -0.11434831;
      W_f[15,18] := 0.06204842;
      W_f[15,19] := -0.16308638;
      W_f[15,20] := -0.08014372;
      W_f[15,21] := 0.09970582;
      W_f[15,22] := -0.01455338;
      W_f[15,23] := -0.09048357;
      W_f[15,24] := 1.48085737;
      W_f[15,25] := 1.43709755;
      W_f[15,26] := -0.04126001;
      W_f[15,27] := 0.03295555;
      W_f[15,28] := -0.08897620;
      W_f[15,29] := 0.14969468;
      W_f[15,30] := 0.12863542;
      W_f[15,31] := -0.01891266;
      W_f[15,32] := -0.08377147;
      W_f[15,33] := 0.04984247;
      W_f[15,34] := 0.73210019;
      W_f[15,35] := -0.07470711;
      W_f[15,36] := 0.01260767;
      W_f[15,37] := -0.02138078;
      W_f[15,38] := 0.01280809;
      W_f[15,39] := 0.12110989;
      W_g[0,0] := 0.13204537;
      W_g[0,1] := -0.07179091;
      W_g[0,2] := 0.13041292;
      W_g[0,3] := -0.01710966;
      W_g[0,4] := 0.08717188;
      W_g[0,5] := -0.03005558;
      W_g[0,6] := 0.02608494;
      W_g[0,7] := -0.02178418;
      W_g[0,8] := -0.02002059;
      W_g[0,9] := -0.01907159;
      W_g[0,10] := -0.07584066;
      W_g[0,11] := -0.02761280;
      W_g[0,12] := -0.03857584;
      W_g[0,13] := -0.01737243;
      W_g[0,14] := -0.10338410;
      W_g[0,15] := -0.00566125;
      W_g[0,16] := -0.01846444;
      W_g[0,17] := -0.09568264;
      W_g[0,18] := 0.01344434;
      W_g[0,19] := -0.04545733;
      W_g[0,20] := -0.07012872;
      W_g[0,21] := -0.22657579;
      W_g[0,22] := -0.00134380;
      W_g[0,23] := 0.01402790;
      W_g[0,24] := 0.05787951;
      W_g[0,25] := 0.33322844;
      W_g[0,26] := 0.13387449;
      W_g[0,27] := -0.28495404;
      W_g[0,28] := 0.08640742;
      W_g[0,29] := 0.00553245;
      W_g[0,30] := 0.00379307;
      W_g[0,31] := 0.00939364;
      W_g[0,32] := -0.02259280;
      W_g[0,33] := -0.03415785;
      W_g[0,34] := 0.41566586;
      W_g[0,35] := -0.02096383;
      W_g[0,36] := -0.04175030;
      W_g[0,37] := -0.04161927;
      W_g[0,38] := 0.04176929;
      W_g[0,39] := -0.02666814;
      W_g[1,0] := 0.10034030;
      W_g[1,1] := 0.02818905;
      W_g[1,2] := 0.08966444;
      W_g[1,3] := 0.02384869;
      W_g[1,4] := -0.00957148;
      W_g[1,5] := 0.02258740;
      W_g[1,6] := 0.21898407;
      W_g[1,7] := 0.03297459;
      W_g[1,8] := 0.02741309;
      W_g[1,9] := 0.03524271;
      W_g[1,10] := -0.09459055;
      W_g[1,11] := 0.00226336;
      W_g[1,12] := -0.03214818;
      W_g[1,13] := 0.09925831;
      W_g[1,14] := 0.03271784;
      W_g[1,15] := -0.00993501;
      W_g[1,16] := 0.04625125;
      W_g[1,17] := -0.01382133;
      W_g[1,18] := 0.14169702;
      W_g[1,19] := -0.06103647;
      W_g[1,20] := -0.21253440;
      W_g[1,21] := 0.11839490;
      W_g[1,22] := -0.01691977;
      W_g[1,23] := 0.05358729;
      W_g[1,24] := -0.32853305;
      W_g[1,25] := -0.49424851;
      W_g[1,26] := -0.08112237;
      W_g[1,27] := 0.12497368;
      W_g[1,28] := 0.17492743;
      W_g[1,29] := 0.05923015;
      W_g[1,30] := -0.03070631;
      W_g[1,31] := -0.01609530;
      W_g[1,32] := 0.01282620;
      W_g[1,33] := 0.00597268;
      W_g[1,34] := -0.44541347;
      W_g[1,35] := 0.04373179;
      W_g[1,36] := 0.07117015;
      W_g[1,37] := -0.05477969;
      W_g[1,38] := -0.11489128;
      W_g[1,39] := -0.05603904;
      W_g[2,0] := -0.03656583;
      W_g[2,1] := 0.08601304;
      W_g[2,2] := -0.02144271;
      W_g[2,3] := -0.00415884;
      W_g[2,4] := 0.05374509;
      W_g[2,5] := 0.01513857;
      W_g[2,6] := 0.00031003;
      W_g[2,7] := -0.00429267;
      W_g[2,8] := 0.00247940;
      W_g[2,9] := -0.02802207;
      W_g[2,10] := 0.00567887;
      W_g[2,11] := 0.07285577;
      W_g[2,12] := 0.06949551;
      W_g[2,13] := -0.06609099;
      W_g[2,14] := 0.02675425;
      W_g[2,15] := 0.05979875;
      W_g[2,16] := 0.18823372;
      W_g[2,17] := 0.10135632;
      W_g[2,18] := -0.01730143;
      W_g[2,19] := 0.07176489;
      W_g[2,20] := -0.00487325;
      W_g[2,21] := -0.01244247;
      W_g[2,22] := 0.07138075;
      W_g[2,23] := -0.08855219;
      W_g[2,24] := 0.66917461;
      W_g[2,25] := 0.40664709;
      W_g[2,26] := 0.05317146;
      W_g[2,27] := -0.03753066;
      W_g[2,28] := 0.04217075;
      W_g[2,29] := -0.08696262;
      W_g[2,30] := 0.07279130;
      W_g[2,31] := 0.04612178;
      W_g[2,32] := 0.06409022;
      W_g[2,33] := 0.01605693;
      W_g[2,34] := 0.15648539;
      W_g[2,35] := 0.11777368;
      W_g[2,36] := -0.03577918;
      W_g[2,37] := -0.02626175;
      W_g[2,38] := -0.29250881;
      W_g[2,39] := -0.17305109;
      W_g[3,0] := 0.03535830;
      W_g[3,1] := -0.10494116;
      W_g[3,2] := 0.03618518;
      W_g[3,3] := -0.03134191;
      W_g[3,4] := -0.24614213;
      W_g[3,5] := 0.12662181;
      W_g[3,6] := 0.06337537;
      W_g[3,7] := -0.03527300;
      W_g[3,8] := -0.03651504;
      W_g[3,9] := -0.03074392;
      W_g[3,10] := -0.05727396;
      W_g[3,11] := -0.02935094;
      W_g[3,12] := -0.03621458;
      W_g[3,13] := -0.01833671;
      W_g[3,14] := -0.16850124;
      W_g[3,15] := -0.00882464;
      W_g[3,16] := -0.02389451;
      W_g[3,17] := -0.07828564;
      W_g[3,18] := 0.02588245;
      W_g[3,19] := -0.04996347;
      W_g[3,20] := -0.03450434;
      W_g[3,21] := 0.08713186;
      W_g[3,22] := 0.04250673;
      W_g[3,23] := 0.02315470;
      W_g[3,24] := 0.24060252;
      W_g[3,25] := -0.04010823;
      W_g[3,26] := -0.04215078;
      W_g[3,27] := 0.04264580;
      W_g[3,28] := -0.24964345;
      W_g[3,29] := -0.01958500;
      W_g[3,30] := 0.03981116;
      W_g[3,31] := 0.05331163;
      W_g[3,32] := 0.02955173;
      W_g[3,33] := 0.03688915;
      W_g[3,34] := -0.07779746;
      W_g[3,35] := 0.04131736;
      W_g[3,36] := -0.09415401;
      W_g[3,37] := 0.02781735;
      W_g[3,38] := -0.01530841;
      W_g[3,39] := -0.10393603;
      W_g[4,0] := 0.07740436;
      W_g[4,1] := -0.07530216;
      W_g[4,2] := 0.08100316;
      W_g[4,3] := -0.03866265;
      W_g[4,4] := -0.12411599;
      W_g[4,5] := -0.06374057;
      W_g[4,6] := -0.06540763;
      W_g[4,7] := -0.05087971;
      W_g[4,8] := -0.02486523;
      W_g[4,9] := -0.00432705;
      W_g[4,10] := -0.02001161;
      W_g[4,11] := -0.22602051;
      W_g[4,12] := -0.27104041;
      W_g[4,13] := -0.04622217;
      W_g[4,14] := 0.03693646;
      W_g[4,15] := -0.22289379;
      W_g[4,16] := -0.03339233;
      W_g[4,17] := -0.10395480;
      W_g[4,18] := -0.67769754;
      W_g[4,19] := -0.10701112;
      W_g[4,20] := -0.00507321;
      W_g[4,21] := 0.06153874;
      W_g[4,22] := -0.05829039;
      W_g[4,23] := -0.03399877;
      W_g[4,24] := 0.02580869;
      W_g[4,25] := -0.05605169;
      W_g[4,26] := 0.02870816;
      W_g[4,27] := 0.09912029;
      W_g[4,28] := -0.08475526;
      W_g[4,29] := 0.02515182;
      W_g[4,30] := -0.06613169;
      W_g[4,31] := -0.01619294;
      W_g[4,32] := -0.07978069;
      W_g[4,33] := -0.02161121;
      W_g[4,34] := -0.01309834;
      W_g[4,35] := -0.05835930;
      W_g[4,36] := 0.02740471;
      W_g[4,37] := -0.06427267;
      W_g[4,38] := -0.14359041;
      W_g[4,39] := -0.04779189;
      W_g[5,0] := 0.07845761;
      W_g[5,1] := 0.12291198;
      W_g[5,2] := 0.09020026;
      W_g[5,3] := -0.05951332;
      W_g[5,4] := -0.18635792;
      W_g[5,5] := -0.67060107;
      W_g[5,6] := -0.09371807;
      W_g[5,7] := -0.06248650;
      W_g[5,8] := -0.05328716;
      W_g[5,9] := -0.05699488;
      W_g[5,10] := -0.21003345;
      W_g[5,11] := -0.04094445;
      W_g[5,12] := -0.03951516;
      W_g[5,13] := 0.01896183;
      W_g[5,14] := 0.05772699;
      W_g[5,15] := -0.03484442;
      W_g[5,16] := -0.08915464;
      W_g[5,17] := -0.03359089;
      W_g[5,18] := 0.05330428;
      W_g[5,19] := -0.04913564;
      W_g[5,20] := -0.02437795;
      W_g[5,21] := -0.03660732;
      W_g[5,22] := 0.05388405;
      W_g[5,23] := 0.03580718;
      W_g[5,24] := 0.66795236;
      W_g[5,25] := 0.38463682;
      W_g[5,26] := 0.03221167;
      W_g[5,27] := -0.09449711;
      W_g[5,28] := -0.21332875;
      W_g[5,29] := -0.10703770;
      W_g[5,30] := 0.04866340;
      W_g[5,31] := 0.04555348;
      W_g[5,32] := 0.03119684;
      W_g[5,33] := 0.02472051;
      W_g[5,34] := -0.00109696;
      W_g[5,35] := 0.00976827;
      W_g[5,36] := -0.04086661;
      W_g[5,37] := 0.01402589;
      W_g[5,38] := 0.01088466;
      W_g[5,39] := 0.05395384;
      W_g[6,0] := -0.09459254;
      W_g[6,1] := -0.34658876;
      W_g[6,2] := -0.12041241;
      W_g[6,3] := 0.11314632;
      W_g[6,4] := 0.07203985;
      W_g[6,5] := -0.09553758;
      W_g[6,6] := -0.03457065;
      W_g[6,7] := 0.12589408;
      W_g[6,8] := 0.09656766;
      W_g[6,9] := 0.12055878;
      W_g[6,10] := 0.01646312;
      W_g[6,11] := -0.06715041;
      W_g[6,12] := -0.08268934;
      W_g[6,13] := -0.01733059;
      W_g[6,14] := 0.05910295;
      W_g[6,15] := -0.07129493;
      W_g[6,16] := -0.06239159;
      W_g[6,17] := -0.06886618;
      W_g[6,18] := 0.04810062;
      W_g[6,19] := -0.09653840;
      W_g[6,20] := 0.16959167;
      W_g[6,21] := -0.00798076;
      W_g[6,22] := 0.00821575;
      W_g[6,23] := 0.10493567;
      W_g[6,24] := 0.06085224;
      W_g[6,25] := 0.05369381;
      W_g[6,26] := -0.02010110;
      W_g[6,27] := 0.00523888;
      W_g[6,28] := -0.05049808;
      W_g[6,29] := 0.04111513;
      W_g[6,30] := 0.01227053;
      W_g[6,31] := 0.02041260;
      W_g[6,32] := -0.00532885;
      W_g[6,33] := -0.00633689;
      W_g[6,34] := -0.01163891;
      W_g[6,35] := 0.03265250;
      W_g[6,36] := -0.08721739;
      W_g[6,37] := 0.02508505;
      W_g[6,38] := -0.13942142;
      W_g[6,39] := -0.03058173;
      W_g[7,0] := 0.13290332;
      W_g[7,1] := -0.22788383;
      W_g[7,2] := 0.14421831;
      W_g[7,3] := -0.04011448;
      W_g[7,4] := -0.00983350;
      W_g[7,5] := 0.06002469;
      W_g[7,6] := 0.01148172;
      W_g[7,7] := -0.03318439;
      W_g[7,8] := -0.04474748;
      W_g[7,9] := -0.03664961;
      W_g[7,10] := -0.05171043;
      W_g[7,11] := 0.15889420;
      W_g[7,12] := 0.18816991;
      W_g[7,13] := 0.03320323;
      W_g[7,14] := 0.08849441;
      W_g[7,15] := 0.10898419;
      W_g[7,16] := -0.10423554;
      W_g[7,17] := 0.21788061;
      W_g[7,18] := -0.09352972;
      W_g[7,19] := 0.22861433;
      W_g[7,20] := 0.01804306;
      W_g[7,21] := 0.02883035;
      W_g[7,22] := 0.02334912;
      W_g[7,23] := 0.00972550;
      W_g[7,24] := 0.09000973;
      W_g[7,25] := 0.23796630;
      W_g[7,26] := -0.00529223;
      W_g[7,27] := 0.02389492;
      W_g[7,28] := 0.01771568;
      W_g[7,29] := 0.03995743;
      W_g[7,30] := 0.02374280;
      W_g[7,31] := 0.00652028;
      W_g[7,32] := 0.02379220;
      W_g[7,33] := 0.01227521;
      W_g[7,34] := -0.02105843;
      W_g[7,35] := 0.02154919;
      W_g[7,36] := -0.01575272;
      W_g[7,37] := -0.01810107;
      W_g[7,38] := -0.00772995;
      W_g[7,39] := -0.28201035;
      W_g[8,0] := 0.01713815;
      W_g[8,1] := -0.00229361;
      W_g[8,2] := 0.01726119;
      W_g[8,3] := -0.02061658;
      W_g[8,4] := -0.04641379;
      W_g[8,5] := 0.04689364;
      W_g[8,6] := 0.00514349;
      W_g[8,7] := -0.02527735;
      W_g[8,8] := -0.02019661;
      W_g[8,9] := -0.01965989;
      W_g[8,10] := -0.02106753;
      W_g[8,11] := -0.18108463;
      W_g[8,12] := -0.17477527;
      W_g[8,13] := -0.07262667;
      W_g[8,14] := 0.09604074;
      W_g[8,15] := -0.22339889;
      W_g[8,16] := -0.01457437;
      W_g[8,17] := 0.18952110;
      W_g[8,18] := 0.09061687;
      W_g[8,19] := -0.16597474;
      W_g[8,20] := -0.02462232;
      W_g[8,21] := -0.08115550;
      W_g[8,22] := 0.02058986;
      W_g[8,23] := -0.05404805;
      W_g[8,24] := -0.07197467;
      W_g[8,25] := -0.24299450;
      W_g[8,26] := 0.03455175;
      W_g[8,27] := -0.12814535;
      W_g[8,28] := -0.12446780;
      W_g[8,29] := -0.07076260;
      W_g[8,30] := 0.03440274;
      W_g[8,31] := 0.02760479;
      W_g[8,32] := -0.00320816;
      W_g[8,33] := -0.00195394;
      W_g[8,34] := -0.06706773;
      W_g[8,35] := -0.03631235;
      W_g[8,36] := -0.04615070;
      W_g[8,37] := 0.02211455;
      W_g[8,38] := 0.00710197;
      W_g[8,39] := 0.06994114;
      W_g[9,0] := -0.26859412;
      W_g[9,1] := -0.16339006;
      W_g[9,2] := -0.30892456;
      W_g[9,3] := -0.12821960;
      W_g[9,4] := 0.01028809;
      W_g[9,5] := -0.05689346;
      W_g[9,6] := 0.13176501;
      W_g[9,7] := -0.11366676;
      W_g[9,8] := -0.13505223;
      W_g[9,9] := -0.13410461;
      W_g[9,10] := -0.29736590;
      W_g[9,11] := 0.03893382;
      W_g[9,12] := 0.03934914;
      W_g[9,13] := 0.01418684;
      W_g[9,14] := 0.01693503;
      W_g[9,15] := 0.04444136;
      W_g[9,16] := 0.07951424;
      W_g[9,17] := 0.00626671;
      W_g[9,18] := -0.06104251;
      W_g[9,19] := 0.04594292;
      W_g[9,20] := -0.02836513;
      W_g[9,21] := 0.03974990;
      W_g[9,22] := -0.02700124;
      W_g[9,23] := 0.02002714;
      W_g[9,24] := -0.50772762;
      W_g[9,25] := -0.25462687;
      W_g[9,26] := -0.03511217;
      W_g[9,27] := 0.04529352;
      W_g[9,28] := 0.04820129;
      W_g[9,29] := 0.09988645;
      W_g[9,30] := -0.01425081;
      W_g[9,31] := -0.01030078;
      W_g[9,32] := -0.01629252;
      W_g[9,33] := -0.00994037;
      W_g[9,34] := -0.59423113;
      W_g[9,35] := 0.03158842;
      W_g[9,36] := -0.08265782;
      W_g[9,37] := -0.03526440;
      W_g[9,38] := -0.00322891;
      W_g[9,39] := -0.00800959;
      W_g[10,0] := -0.03213325;
      W_g[10,1] := -0.00863164;
      W_g[10,2] := -0.03062097;
      W_g[10,3] := 0.01255380;
      W_g[10,4] := 0.10173590;
      W_g[10,5] := -0.04505892;
      W_g[10,6] := -0.00103756;
      W_g[10,7] := 0.01735601;
      W_g[10,8] := 0.01301922;
      W_g[10,9] := 0.01365640;
      W_g[10,10] := 0.00548952;
      W_g[10,11] := -0.00245858;
      W_g[10,12] := 0.00857112;
      W_g[10,13] := 0.10749885;
      W_g[10,14] := -0.12755091;
      W_g[10,15] := -0.03629598;
      W_g[10,16] := -0.01334849;
      W_g[10,17] := 0.12906626;
      W_g[10,18] := -0.01503343;
      W_g[10,19] := 0.01173486;
      W_g[10,20] := 0.06222534;
      W_g[10,21] := 0.05678142;
      W_g[10,22] := -0.02349397;
      W_g[10,23] := 0.06754656;
      W_g[10,24] := 0.17796169;
      W_g[10,25] := 0.19162965;
      W_g[10,26] := -0.02255434;
      W_g[10,27] := 0.10073226;
      W_g[10,28] := 0.13280237;
      W_g[10,29] := -0.01282987;
      W_g[10,30] := -0.01621767;
      W_g[10,31] := -0.01406650;
      W_g[10,32] := -0.00099214;
      W_g[10,33] := -0.00035058;
      W_g[10,34] := 0.14521876;
      W_g[10,35] := 0.02793738;
      W_g[10,36] := -0.07625148;
      W_g[10,37] := -0.00763791;
      W_g[10,38] := 0.00534324;
      W_g[10,39] := -0.33125421;
      W_g[11,0] := -0.11375076;
      W_g[11,1] := 0.05398307;
      W_g[11,2] := -0.12075092;
      W_g[11,3] := 0.04525032;
      W_g[11,4] := 0.08992387;
      W_g[11,5] := 0.01991016;
      W_g[11,6] := 0.22497544;
      W_g[11,7] := 0.04191377;
      W_g[11,8] := 0.04533296;
      W_g[11,9] := 0.04499990;
      W_g[11,10] := -0.10994546;
      W_g[11,11] := 0.00437518;
      W_g[11,12] := -0.00140931;
      W_g[11,13] := 0.04130397;
      W_g[11,14] := 0.05369400;
      W_g[11,15] := -0.00366092;
      W_g[11,16] := -0.07105832;
      W_g[11,17] := -0.07482163;
      W_g[11,18] := -0.07100122;
      W_g[11,19] := 0.01718117;
      W_g[11,20] := -0.13757822;
      W_g[11,21] := 0.11307504;
      W_g[11,22] := 0.05416900;
      W_g[11,23] := 0.02884634;
      W_g[11,24] := 0.53078175;
      W_g[11,25] := 0.35704109;
      W_g[11,26] := 0.03378000;
      W_g[11,27] := 0.10375553;
      W_g[11,28] := 0.25050017;
      W_g[11,29] := -0.12446285;
      W_g[11,30] := 0.05581930;
      W_g[11,31] := 0.05851344;
      W_g[11,32] := 0.07730477;
      W_g[11,33] := 0.09541148;
      W_g[11,34] := 0.12033152;
      W_g[11,35] := 0.12105432;
      W_g[11,36] := -0.19497558;
      W_g[11,37] := 0.01371960;
      W_g[11,38] := 0.08832928;
      W_g[11,39] := 0.08146589;
      W_g[12,0] := -0.02631861;
      W_g[12,1] := 0.04126604;
      W_g[12,2] := -0.02663527;
      W_g[12,3] := -0.02984582;
      W_g[12,4] := -0.02636349;
      W_g[12,5] := 0.07986053;
      W_g[12,6] := -0.01390989;
      W_g[12,7] := -0.00909171;
      W_g[12,8] := -0.01941176;
      W_g[12,9] := -0.02868326;
      W_g[12,10] := 0.03089914;
      W_g[12,11] := 0.00787742;
      W_g[12,12] := -0.00904082;
      W_g[12,13] := -0.02910480;
      W_g[12,14] := 0.10839512;
      W_g[12,15] := 0.01380038;
      W_g[12,16] := 0.06520407;
      W_g[12,17] := -0.04494612;
      W_g[12,18] := -0.00194090;
      W_g[12,19] := -0.01509680;
      W_g[12,20] := 0.08029543;
      W_g[12,21] := 0.02437602;
      W_g[12,22] := -0.07042312;
      W_g[12,23] := -0.04948704;
      W_g[12,24] := -0.83039939;
      W_g[12,25] := -0.55899370;
      W_g[12,26] := -0.04566456;
      W_g[12,27] := 0.00189110;
      W_g[12,28] := -0.02951618;
      W_g[12,29] := -0.05513477;
      W_g[12,30] := -0.04795056;
      W_g[12,31] := -0.03688380;
      W_g[12,32] := -0.03588131;
      W_g[12,33] := 0.00737297;
      W_g[12,34] := 0.04994570;
      W_g[12,35] := -0.01839683;
      W_g[12,36] := -0.49873567;
      W_g[12,37] := -0.07791845;
      W_g[12,38] := -0.10474910;
      W_g[12,39] := 0.00553967;
      W_g[13,0] := -0.02684040;
      W_g[13,1] := -0.08890500;
      W_g[13,2] := -0.02790045;
      W_g[13,3] := 0.08189317;
      W_g[13,4] := -0.12551519;
      W_g[13,5] := -0.05772218;
      W_g[13,6] := 0.09080454;
      W_g[13,7] := 0.08241173;
      W_g[13,8] := 0.07553043;
      W_g[13,9] := 0.08949121;
      W_g[13,10] := -0.02704351;
      W_g[13,11] := 0.00487661;
      W_g[13,12] := 0.02095871;
      W_g[13,13] := 0.06879441;
      W_g[13,14] := 0.00018557;
      W_g[13,15] := 0.01617457;
      W_g[13,16] := 0.23046753;
      W_g[13,17] := 0.08005539;
      W_g[13,18] := -0.06847396;
      W_g[13,19] := 0.02106568;
      W_g[13,20] := -0.08102658;
      W_g[13,21] := -0.03850572;
      W_g[13,22] := 0.00878646;
      W_g[13,23] := 0.14752086;
      W_g[13,24] := 0.19677557;
      W_g[13,25] := -0.00969006;
      W_g[13,26] := 0.04820746;
      W_g[13,27] := -0.06298333;
      W_g[13,28] := -0.06368192;
      W_g[13,29] := 0.01809042;
      W_g[13,30] := 0.01814866;
      W_g[13,31] := 0.00847225;
      W_g[13,32] := 0.00546922;
      W_g[13,33] := -0.01145526;
      W_g[13,34] := 0.13813621;
      W_g[13,35] := 0.01473064;
      W_g[13,36] := -0.05009100;
      W_g[13,37] := -0.01566363;
      W_g[13,38] := 0.05946118;
      W_g[13,39] := 0.00826691;
      W_g[14,0] := 0.02104861;
      W_g[14,1] := 0.02198478;
      W_g[14,2] := 0.01118620;
      W_g[14,3] := -0.06436396;
      W_g[14,4] := 0.00489476;
      W_g[14,5] := 0.09250024;
      W_g[14,6] := -0.03399736;
      W_g[14,7] := -0.04967630;
      W_g[14,8] := -0.05370576;
      W_g[14,9] := -0.05536002;
      W_g[14,10] := 0.01229766;
      W_g[14,11] := -0.01784988;
      W_g[14,12] := -0.03607991;
      W_g[14,13] := 0.19007476;
      W_g[14,14] := 0.08048796;
      W_g[14,15] := -0.00893450;
      W_g[14,16] := 0.01208448;
      W_g[14,17] := -0.06566814;
      W_g[14,18] := -0.22113875;
      W_g[14,19] := -0.04166633;
      W_g[14,20] := 0.07567322;
      W_g[14,21] := -0.00166608;
      W_g[14,22] := -0.01256561;
      W_g[14,23] := 0.15394352;
      W_g[14,24] := 0.03526039;
      W_g[14,25] := 0.48119587;
      W_g[14,26] := 0.01489335;
      W_g[14,27] := 0.03173870;
      W_g[14,28] := 0.01991428;
      W_g[14,29] := 0.03107417;
      W_g[14,30] := -0.00682632;
      W_g[14,31] := 0.00660902;
      W_g[14,32] := 0.00283587;
      W_g[14,33] := -0.00859028;
      W_g[14,34] := -0.02930867;
      W_g[14,35] := 0.03631073;
      W_g[14,36] := 0.00467363;
      W_g[14,37] := 0.02703222;
      W_g[14,38] := -0.04237745;
      W_g[14,39] := 0.01309555;
      W_g[15,0] := 0.08495549;
      W_g[15,1] := -0.20728092;
      W_g[15,2] := 0.08629236;
      W_g[15,3] := -0.06330224;
      W_g[15,4] := 0.19237527;
      W_g[15,5] := 0.00801008;
      W_g[15,6] := -0.10499398;
      W_g[15,7] := -0.05814644;
      W_g[15,8] := -0.06757385;
      W_g[15,9] := -0.05901760;
      W_g[15,10] := -0.00683508;
      W_g[15,11] := -0.00540838;
      W_g[15,12] := -0.02551957;
      W_g[15,13] := -0.01507952;
      W_g[15,14] := 0.00483655;
      W_g[15,15] := 0.01358667;
      W_g[15,16] := 0.25418368;
      W_g[15,17] := -0.01636837;
      W_g[15,18] := 0.01947031;
      W_g[15,19] := -0.03640394;
      W_g[15,20] := 0.21466117;
      W_g[15,21] := 0.10691275;
      W_g[15,22] := 0.03332973;
      W_g[15,23] := -0.06589723;
      W_g[15,24] := 0.15037987;
      W_g[15,25] := 0.03056319;
      W_g[15,26] := -0.08210966;
      W_g[15,27] := 0.14967138;
      W_g[15,28] := 0.09097399;
      W_g[15,29] := -0.04645663;
      W_g[15,30] := 0.04627259;
      W_g[15,31] := 0.00594573;
      W_g[15,32] := 0.05130993;
      W_g[15,33] := 0.05626767;
      W_g[15,34] := -0.00315162;
      W_g[15,35] := 0.04370028;
      W_g[15,36] := -0.06999733;
      W_g[15,37] := 0.01681984;
      W_g[15,38] := 0.07271070;
      W_g[15,39] := 0.01082875;
      W_o[0,0] := -0.19233570;
      W_o[0,1] := 0.16228242;
      W_o[0,2] := 0.03764162;
      W_o[0,3] := -0.00444271;
      W_o[0,4] := 0.08973370;
      W_o[0,5] := 0.05718408;
      W_o[0,6] := -0.23139432;
      W_o[0,7] := 0.15783574;
      W_o[0,8] := -0.15828826;
      W_o[0,9] := 0.19736247;
      W_o[0,10] := -0.30527124;
      W_o[0,11] := -0.23014921;
      W_o[0,12] := 0.20966798;
      W_o[0,13] := -0.17421527;
      W_o[0,14] := -0.26786944;
      W_o[0,15] := -0.01321167;
      W_o[0,16] := -0.01970488;
      W_o[0,17] := -0.20280616;
      W_o[0,18] := 0.42725509;
      W_o[0,19] := -0.06582518;
      W_o[0,20] := -0.03046696;
      W_o[0,21] := 0.55015820;
      W_o[0,22] := 0.44234657;
      W_o[0,23] := -0.33459106;
      W_o[0,24] := 1.26524746;
      W_o[0,25] := 1.41665208;
      W_o[0,26] := -0.32673731;
      W_o[0,27] := -0.18320346;
      W_o[0,28] := 0.01126313;
      W_o[0,29] := -0.28385833;
      W_o[0,30] := 0.26098812;
      W_o[0,31] := 0.04669111;
      W_o[0,32] := 0.10434872;
      W_o[0,33] := 0.05575988;
      W_o[0,34] := 1.33235300;
      W_o[0,35] := -0.06145113;
      W_o[0,36] := -0.03345130;
      W_o[0,37] := -0.22215474;
      W_o[0,38] := 0.00487359;
      W_o[0,39] := -0.03890218;
      W_o[1,0] := 0.74378037;
      W_o[1,1] := -0.05000130;
      W_o[1,2] := 0.12129822;
      W_o[1,3] := 0.10320133;
      W_o[1,4] := 0.11998425;
      W_o[1,5] := -0.19072209;
      W_o[1,6] := 0.21001612;
      W_o[1,7] := 0.11332466;
      W_o[1,8] := 0.35882619;
      W_o[1,9] := 0.38575748;
      W_o[1,10] := -0.45878416;
      W_o[1,11] := -0.15748191;
      W_o[1,12] := 0.20664066;
      W_o[1,13] := 0.12306170;
      W_o[1,14] := -0.20303696;
      W_o[1,15] := 0.03768912;
      W_o[1,16] := -0.05619529;
      W_o[1,17] := -0.09439399;
      W_o[1,18] := 0.27072540;
      W_o[1,19] := 0.38222137;
      W_o[1,20] := -0.29343513;
      W_o[1,21] := 0.51613772;
      W_o[1,22] := 0.17591031;
      W_o[1,23] := 0.18373588;
      W_o[1,24] := -0.03005522;
      W_o[1,25] := 0.00781888;
      W_o[1,26] := -0.10684884;
      W_o[1,27] := -0.07173182;
      W_o[1,28] := 0.20145275;
      W_o[1,29] := 0.13064608;
      W_o[1,30] := -0.01024106;
      W_o[1,31] := -0.07163240;
      W_o[1,32] := 0.05804014;
      W_o[1,33] := 0.27217436;
      W_o[1,34] := 0.06194695;
      W_o[1,35] := -0.30407301;
      W_o[1,36] := 0.15308920;
      W_o[1,37] := -0.07396729;
      W_o[1,38] := 0.08739793;
      W_o[1,39] := 0.32655314;
      W_o[2,0] := -0.03605163;
      W_o[2,1] := 0.07661975;
      W_o[2,2] := 0.13695037;
      W_o[2,3] := 0.09188601;
      W_o[2,4] := 0.03664814;
      W_o[2,5] := -0.02675835;
      W_o[2,6] := -0.01984608;
      W_o[2,7] := -0.19014685;
      W_o[2,8] := -0.02938575;
      W_o[2,9] := 0.18366605;
      W_o[2,10] := -0.18625411;
      W_o[2,11] := 0.06671655;
      W_o[2,12] := 0.31907275;
      W_o[2,13] := -0.01547686;
      W_o[2,14] := -0.05195596;
      W_o[2,15] := 0.03504787;
      W_o[2,16] := 0.35419029;
      W_o[2,17] := 0.02718459;
      W_o[2,18] := -0.24911258;
      W_o[2,19] := -0.86676186;
      W_o[2,20] := -0.12667567;
      W_o[2,21] := 0.02015731;
      W_o[2,22] := -0.02294585;
      W_o[2,23] := -0.01648583;
      W_o[2,24] := -0.19191538;
      W_o[2,25] := 0.00051678;
      W_o[2,26] := 0.06543333;
      W_o[2,27] := 0.10374146;
      W_o[2,28] := -0.04504570;
      W_o[2,29] := 0.21506196;
      W_o[2,30] := 0.02658869;
      W_o[2,31] := -0.13691518;
      W_o[2,32] := 0.01719045;
      W_o[2,33] := 0.21874297;
      W_o[2,34] := -0.07076459;
      W_o[2,35] := -0.07407880;
      W_o[2,36] := -0.08052358;
      W_o[2,37] := -0.20128877;
      W_o[2,38] := -0.38490325;
      W_o[2,39] := 0.68916357;
      W_o[3,0] := -0.06302688;
      W_o[3,1] := 0.20022115;
      W_o[3,2] := 0.01595870;
      W_o[3,3] := -0.00183610;
      W_o[3,4] := -0.85917354;
      W_o[3,5] := 0.17318121;
      W_o[3,6] := 0.24098408;
      W_o[3,7] := 0.25960821;
      W_o[3,8] := -0.00940404;
      W_o[3,9] := 0.06814823;
      W_o[3,10] := -0.01664601;
      W_o[3,11] := 0.14877798;
      W_o[3,12] := -0.09583785;
      W_o[3,13] := -0.27983487;
      W_o[3,14] := 0.14434218;
      W_o[3,15] := 0.00555357;
      W_o[3,16] := -0.02839783;
      W_o[3,17] := 0.09947813;
      W_o[3,18] := 0.46432632;
      W_o[3,19] := 0.06364350;
      W_o[3,20] := -0.08531965;
      W_o[3,21] := 1.16577530;
      W_o[3,22] := 0.34482756;
      W_o[3,23] := -0.11727701;
      W_o[3,24] := 1.35247672;
      W_o[3,25] := 1.17824149;
      W_o[3,26] := -0.48925292;
      W_o[3,27] := -0.77375019;
      W_o[3,28] := 0.22645181;
      W_o[3,29] := 0.00574818;
      W_o[3,30] := 0.24614631;
      W_o[3,31] := 0.10528258;
      W_o[3,32] := 0.00088265;
      W_o[3,33] := 0.10498052;
      W_o[3,34] := 1.18573022;
      W_o[3,35] := 0.19094193;
      W_o[3,36] := -0.00811989;
      W_o[3,37] := 0.09236411;
      W_o[3,38] := 0.11084373;
      W_o[3,39] := 0.92378908;
      W_o[4,0] := -0.18556677;
      W_o[4,1] := -0.06182796;
      W_o[4,2] := 0.14978686;
      W_o[4,3] := -0.02874054;
      W_o[4,4] := -0.23721895;
      W_o[4,5] := -0.02661614;
      W_o[4,6] := 0.04865195;
      W_o[4,7] := -0.25955087;
      W_o[4,8] := 0.51465279;
      W_o[4,9] := -0.28220513;
      W_o[4,10] := 0.01177313;
      W_o[4,11] := -0.49890938;
      W_o[4,12] := -0.86487442;
      W_o[4,13] := -0.04488994;
      W_o[4,14] := -0.05423390;
      W_o[4,15] := -0.55890763;
      W_o[4,16] := -0.14559400;
      W_o[4,17] := 0.02167914;
      W_o[4,18] := 1.00664401;
      W_o[4,19] := -0.25995746;
      W_o[4,20] := 0.00703312;
      W_o[4,21] := -0.22832327;
      W_o[4,22] := 0.00192229;
      W_o[4,23] := -0.01435418;
      W_o[4,24] := 0.04472705;
      W_o[4,25] := 0.23385289;
      W_o[4,26] := -0.11271448;
      W_o[4,27] := 0.08130027;
      W_o[4,28] := 0.46038952;
      W_o[4,29] := 0.13796063;
      W_o[4,30] := 0.18121891;
      W_o[4,31] := -0.39012441;
      W_o[4,32] := -0.07037880;
      W_o[4,33] := 0.28881219;
      W_o[4,34] := 0.40345052;
      W_o[4,35] := 0.03288190;
      W_o[4,36] := -0.09105004;
      W_o[4,37] := 0.09711539;
      W_o[4,38] := -0.19107214;
      W_o[4,39] := -0.01934181;
      W_o[5,0] := -0.65951943;
      W_o[5,1] := 0.37721992;
      W_o[5,2] := 0.00501744;
      W_o[5,3] := 0.53254199;
      W_o[5,4] := 0.23661830;
      W_o[5,5] := 1.09201050;
      W_o[5,6] := 0.95025426;
      W_o[5,7] := 0.25825107;
      W_o[5,8] := -0.46912813;
      W_o[5,9] := 0.39281145;
      W_o[5,10] := 1.11464036;
      W_o[5,11] := -0.77818263;
      W_o[5,12] := -0.60747635;
      W_o[5,13] := 0.16800997;
      W_o[5,14] := -0.10865308;
      W_o[5,15] := -0.68417382;
      W_o[5,16] := -0.36786407;
      W_o[5,17] := -0.21723378;
      W_o[5,18] := 0.38631910;
      W_o[5,19] := -0.49505970;
      W_o[5,20] := -0.51198816;
      W_o[5,21] := -0.17804918;
      W_o[5,22] := 0.15449362;
      W_o[5,23] := 0.13831171;
      W_o[5,24] := 1.00488901;
      W_o[5,25] := 1.13941503;
      W_o[5,26] := -0.30153662;
      W_o[5,27] := -0.04238907;
      W_o[5,28] := -0.31084278;
      W_o[5,29] := 0.39699879;
      W_o[5,30] := 0.01171695;
      W_o[5,31] := -0.31396887;
      W_o[5,32] := -0.32433808;
      W_o[5,33] := -0.41490105;
      W_o[5,34] := 0.22155695;
      W_o[5,35] := -0.13369399;
      W_o[5,36] := 0.02332771;
      W_o[5,37] := -0.14874032;
      W_o[5,38] := 0.19793962;
      W_o[5,39] := -0.20301516;
      W_o[6,0] := -0.04529256;
      W_o[6,1] := 0.21502827;
      W_o[6,2] := 0.09295318;
      W_o[6,3] := -0.07670660;
      W_o[6,4] := -0.12364518;
      W_o[6,5] := 0.35737661;
      W_o[6,6] := -0.26468867;
      W_o[6,7] := 0.28348017;
      W_o[6,8] := -0.04882327;
      W_o[6,9] := 0.84130001;
      W_o[6,10] := 1.08996773;
      W_o[6,11] := -0.06981075;
      W_o[6,12] := 0.05921048;
      W_o[6,13] := -0.50993186;
      W_o[6,14] := 0.04131682;
      W_o[6,15] := 0.09513918;
      W_o[6,16] := 0.08072844;
      W_o[6,17] := 0.02096614;
      W_o[6,18] := 0.16838115;
      W_o[6,19] := 0.11047240;
      W_o[6,20] := -0.33922145;
      W_o[6,21] := -0.09979945;
      W_o[6,22] := 0.15019019;
      W_o[6,23] := -0.06504018;
      W_o[6,24] := 1.94938886;
      W_o[6,25] := 1.97998226;
      W_o[6,26] := 0.02307883;
      W_o[6,27] := 0.26848882;
      W_o[6,28] := 0.09674384;
      W_o[6,29] := 0.21163414;
      W_o[6,30] := 0.14136782;
      W_o[6,31] := -0.01244890;
      W_o[6,32] := -0.04519035;
      W_o[6,33] := -0.13967720;
      W_o[6,34] := 0.49392059;
      W_o[6,35] := -0.21307352;
      W_o[6,36] := 0.06053885;
      W_o[6,37] := 0.05874070;
      W_o[6,38] := 0.42970201;
      W_o[6,39] := -0.10621832;
      W_o[7,0] := 0.16481332;
      W_o[7,1] := -0.09838933;
      W_o[7,2] := -0.09392150;
      W_o[7,3] := -0.12725453;
      W_o[7,4] := -0.23335472;
      W_o[7,5] := 0.05955706;
      W_o[7,6] := 0.27170953;
      W_o[7,7] := 0.11008973;
      W_o[7,8] := 0.18096824;
      W_o[7,9] := 0.01596895;
      W_o[7,10] := 0.14986110;
      W_o[7,11] := -0.31007567;
      W_o[7,12] := 0.53089291;
      W_o[7,13] := -0.07378945;
      W_o[7,14] := -0.25098050;
      W_o[7,15] := 0.26493293;
      W_o[7,16] := -0.14761060;
      W_o[7,17] := -0.23922910;
      W_o[7,18] := 0.40801761;
      W_o[7,19] := -0.15047765;
      W_o[7,20] := -0.11114324;
      W_o[7,21] := 0.11321358;
      W_o[7,22] := 0.46452600;
      W_o[7,23] := -0.13142034;
      W_o[7,24] := 0.85248584;
      W_o[7,25] := 0.93194580;
      W_o[7,26] := 0.19103780;
      W_o[7,27] := -0.04179411;
      W_o[7,28] := 0.17278184;
      W_o[7,29] := -0.34189469;
      W_o[7,30] := 0.47304693;
      W_o[7,31] := 0.08789608;
      W_o[7,32] := 0.21707091;
      W_o[7,33] := -0.03279238;
      W_o[7,34] := 0.65826845;
      W_o[7,35] := 0.08038806;
      W_o[7,36] := 0.04812925;
      W_o[7,37] := 0.43783510;
      W_o[7,38] := -0.06570955;
      W_o[7,39] := -1.68170238;
      W_o[8,0] := 0.28385592;
      W_o[8,1] := -0.13761093;
      W_o[8,2] := -0.00303996;
      W_o[8,3] := -0.15149458;
      W_o[8,4] := -0.05367951;
      W_o[8,5] := 0.37584558;
      W_o[8,6] := 0.02626968;
      W_o[8,7] := -0.14221786;
      W_o[8,8] := 0.00944922;
      W_o[8,9] := -0.20793188;
      W_o[8,10] := -0.21312512;
      W_o[8,11] := -1.02598393;
      W_o[8,12] := -0.39852768;
      W_o[8,13] := -0.08186030;
      W_o[8,14] := -0.10520020;
      W_o[8,15] := -1.12057710;
      W_o[8,16] := 0.05219958;
      W_o[8,17] := 0.79091048;
      W_o[8,18] := 0.37796351;
      W_o[8,19] := 0.16328999;
      W_o[8,20] := -0.06752818;
      W_o[8,21] := 0.22449610;
      W_o[8,22] := -0.13329799;
      W_o[8,23] := -0.54986066;
      W_o[8,24] := 0.21067502;
      W_o[8,25] := 0.42498264;
      W_o[8,26] := 0.30855075;
      W_o[8,27] := 0.00327513;
      W_o[8,28] := -0.13286735;
      W_o[8,29] := 0.24233432;
      W_o[8,30] := -0.29167452;
      W_o[8,31] := 0.11131452;
      W_o[8,32] := 0.23540798;
      W_o[8,33] := 0.25938869;
      W_o[8,34] := 0.26193738;
      W_o[8,35] := 0.09260385;
      W_o[8,36] := -0.07284077;
      W_o[8,37] := 0.27167174;
      W_o[8,38] := -0.59216839;
      W_o[8,39] := 0.16132931;
      W_o[9,0] := -0.63450861;
      W_o[9,1] := -0.25937200;
      W_o[9,2] := -0.44104776;
      W_o[9,3] := -0.14795317;
      W_o[9,4] := 0.07470662;
      W_o[9,5] := -0.14423917;
      W_o[9,6] := 0.20446719;
      W_o[9,7] := -0.36297330;
      W_o[9,8] := -0.83572245;
      W_o[9,9] := -0.03687909;
      W_o[9,10] := -0.52778012;
      W_o[9,11] := 0.13956045;
      W_o[9,12] := 0.00705423;
      W_o[9,13] := -0.06065191;
      W_o[9,14] := 0.00270301;
      W_o[9,15] := 0.02473978;
      W_o[9,16] := -0.13662922;
      W_o[9,17] := -0.11914370;
      W_o[9,18] := -0.06459489;
      W_o[9,19] := -0.15596199;
      W_o[9,20] := -0.13322008;
      W_o[9,21] := 0.61681378;
      W_o[9,22] := -0.00820900;
      W_o[9,23] := -0.03221058;
      W_o[9,24] := -0.07914114;
      W_o[9,25] := -0.28223765;
      W_o[9,26] := 0.17991577;
      W_o[9,27] := 0.13542831;
      W_o[9,28] := 0.19057170;
      W_o[9,29] := 0.32574418;
      W_o[9,30] := 0.20454229;
      W_o[9,31] := 0.11754695;
      W_o[9,32] := 0.18692589;
      W_o[9,33] := 0.41695151;
      W_o[9,34] := 0.13182598;
      W_o[9,35] := -0.18678822;
      W_o[9,36] := -0.09728058;
      W_o[9,37] := -0.21517648;
      W_o[9,38] := 0.03850761;
      W_o[9,39] := -0.00446410;
      W_o[10,0] := 0.06105608;
      W_o[10,1] := -0.06832715;
      W_o[10,2] := 0.07474305;
      W_o[10,3] := -0.08913961;
      W_o[10,4] := -0.23275980;
      W_o[10,5] := 0.07582341;
      W_o[10,6] := 0.10436798;
      W_o[10,7] := 0.03688281;
      W_o[10,8] := -0.01102509;
      W_o[10,9] := -0.02805536;
      W_o[10,10] := 0.10925468;
      W_o[10,11] := -0.04491638;
      W_o[10,12] := -0.00955069;
      W_o[10,13] := -0.36002284;
      W_o[10,14] := -0.25981170;
      W_o[10,15] := -0.13129516;
      W_o[10,16] := 0.12702818;
      W_o[10,17] := 0.24559321;
      W_o[10,18] := 0.02347365;
      W_o[10,19] := 0.08953306;
      W_o[10,20] := -0.41282898;
      W_o[10,21] := -0.12692606;
      W_o[10,22] := 0.14309493;
      W_o[10,23] := -0.28836918;
      W_o[10,24] := 1.61310303;
      W_o[10,25] := 1.56905019;
      W_o[10,26] := 0.11707000;
      W_o[10,27] := -0.62532181;
      W_o[10,28] := -0.57065505;
      W_o[10,29] := 0.06348585;
      W_o[10,30] := 0.21993062;
      W_o[10,31] := -0.02762064;
      W_o[10,32] := 0.08508236;
      W_o[10,33] := 0.26037309;
      W_o[10,34] := 0.52386832;
      W_o[10,35] := -0.30729154;
      W_o[10,36] := 0.45898029;
      W_o[10,37] := -0.32611471;
      W_o[10,38] := -0.04951124;
      W_o[10,39] := -0.01655830;
      W_o[11,0] := 0.27178949;
      W_o[11,1] := 0.49731860;
      W_o[11,2] := -0.11114703;
      W_o[11,3] := 0.00516717;
      W_o[11,4] := -0.72877467;
      W_o[11,5] := -0.07876529;
      W_o[11,6] := -0.50726026;
      W_o[11,7] := -0.03536538;
      W_o[11,8] := 0.12013210;
      W_o[11,9] := 0.11127870;
      W_o[11,10] := 0.15323649;
      W_o[11,11] := -0.48916084;
      W_o[11,12] := 0.18876550;
      W_o[11,13] := 0.18523493;
      W_o[11,14] := 0.17033486;
      W_o[11,15] := -0.24672720;
      W_o[11,16] := 0.04845995;
      W_o[11,17] := 0.28191727;
      W_o[11,18] := 0.10573061;
      W_o[11,19] := -0.00306271;
      W_o[11,20] := -0.72405404;
      W_o[11,21] := 0.09254762;
      W_o[11,22] := -0.40998662;
      W_o[11,23] := -0.10736269;
      W_o[11,24] := -0.05867720;
      W_o[11,25] := 0.34301037;
      W_o[11,26] := 0.18553430;
      W_o[11,27] := 0.10847312;
      W_o[11,28] := 0.50402117;
      W_o[11,29] := -0.00853192;
      W_o[11,30] := -0.36624411;
      W_o[11,31] := -0.01966033;
      W_o[11,32] := -0.06275205;
      W_o[11,33] := 0.09751767;
      W_o[11,34] := -0.20046946;
      W_o[11,35] := -0.10344042;
      W_o[11,36] := 0.23024116;
      W_o[11,37] := 0.14145058;
      W_o[11,38] := 0.26650199;
      W_o[11,39] := -0.30978867;
      W_o[12,0] := -0.01830707;
      W_o[12,1] := 0.13116099;
      W_o[12,2] := 0.00496979;
      W_o[12,3] := 0.20619306;
      W_o[12,4] := 0.03057155;
      W_o[12,5] := 0.02297443;
      W_o[12,6] := 0.05931674;
      W_o[12,7] := -0.03210922;
      W_o[12,8] := 0.07573608;
      W_o[12,9] := 0.12480564;
      W_o[12,10] := -0.07253183;
      W_o[12,11] := -0.24422289;
      W_o[12,12] := 0.13263887;
      W_o[12,13] := -0.16643250;
      W_o[12,14] := -0.14052729;
      W_o[12,15] := -0.05658006;
      W_o[12,16] := 0.04406866;
      W_o[12,17] := 0.02368420;
      W_o[12,18] := 0.79103941;
      W_o[12,19] := 0.02559086;
      W_o[12,20] := -0.16355352;
      W_o[12,21] := -0.01013497;
      W_o[12,22] := -0.35066113;
      W_o[12,23] := -0.18857741;
      W_o[12,24] := 0.49971122;
      W_o[12,25] := 0.51548553;
      W_o[12,26] := 0.18439379;
      W_o[12,27] := 0.02656424;
      W_o[12,28] := 0.00674596;
      W_o[12,29] := 0.03458697;
      W_o[12,30] := -0.43187174;
      W_o[12,31] := -0.13124835;
      W_o[12,32] := -0.38121006;
      W_o[12,33] := -0.02800291;
      W_o[12,34] := -0.22859025;
      W_o[12,35] := 0.12376902;
      W_o[12,36] := 0.08067092;
      W_o[12,37] := -0.04127869;
      W_o[12,38] := -0.06010977;
      W_o[12,39] := -0.00181283;
      W_o[13,0] := -0.04045204;
      W_o[13,1] := -0.39684391;
      W_o[13,2] := 0.08165251;
      W_o[13,3] := -0.01278869;
      W_o[13,4] := -0.44792256;
      W_o[13,5] := -0.26560831;
      W_o[13,6] := 0.32351243;
      W_o[13,7] := 0.57420599;
      W_o[13,8] := -0.27941430;
      W_o[13,9] := 0.35983771;
      W_o[13,10] := -0.08126416;
      W_o[13,11] := -0.00919488;
      W_o[13,12] := 0.09122144;
      W_o[13,13] := 0.02155786;
      W_o[13,14] := 0.12092461;
      W_o[13,15] := -0.00289959;
      W_o[13,16] := -0.25493520;
      W_o[13,17] := -0.24869688;
      W_o[13,18] := 0.69173944;
      W_o[13,19] := -0.03206153;
      W_o[13,20] := -0.22193044;
      W_o[13,21] := 0.11834586;
      W_o[13,22] := 0.36793059;
      W_o[13,23] := 0.44132417;
      W_o[13,24] := 1.97520661;
      W_o[13,25] := 1.84376884;
      W_o[13,26] := -0.27926096;
      W_o[13,27] := -0.30778426;
      W_o[13,28] := -0.01960251;
      W_o[13,29] := -0.23696770;
      W_o[13,30] := 0.10964504;
      W_o[13,31] := -0.10797819;
      W_o[13,32] := 0.03879900;
      W_o[13,33] := 0.05485996;
      W_o[13,34] := 0.59725481;
      W_o[13,35] := 0.01886969;
      W_o[13,36] := 0.09835773;
      W_o[13,37] := 0.38435343;
      W_o[13,38] := 0.05617079;
      W_o[13,39] := -0.22277038;
      W_o[14,0] := 0.82890773;
      W_o[14,1] := -0.20311049;
      W_o[14,2] := 0.03403382;
      W_o[14,3] := 0.05452057;
      W_o[14,4] := 0.22728330;
      W_o[14,5] := -0.07046781;
      W_o[14,6] := 0.38965160;
      W_o[14,7] := 0.48719046;
      W_o[14,8] := -0.07724485;
      W_o[14,9] := -0.07247894;
      W_o[14,10] := 0.28147829;
      W_o[14,11] := -0.02350411;
      W_o[14,12] := 0.37411377;
      W_o[14,13] := 0.01457606;
      W_o[14,14] := -0.08907567;
      W_o[14,15] := 0.03109477;
      W_o[14,16] := 0.05151353;
      W_o[14,17] := -0.15667544;
      W_o[14,18] := -0.26403114;
      W_o[14,19] := -0.10761543;
      W_o[14,20] := 0.38541514;
      W_o[14,21] := 1.57582223;
      W_o[14,22] := -0.05344179;
      W_o[14,23] := -0.94024462;
      W_o[14,24] := -0.01890260;
      W_o[14,25] := -0.00721721;
      W_o[14,26] := -0.42063591;
      W_o[14,27] := 0.50790477;
      W_o[14,28] := 0.23005128;
      W_o[14,29] := 0.23416848;
      W_o[14,30] := -0.10726156;
      W_o[14,31] := -0.05015407;
      W_o[14,32] := 0.03626099;
      W_o[14,33] := 0.22095527;
      W_o[14,34] := 0.28296489;
      W_o[14,35] := -0.10200696;
      W_o[14,36] := 0.00415739;
      W_o[14,37] := 0.20215775;
      W_o[14,38] := 0.14493252;
      W_o[14,39] := 0.19539395;
      W_o[15,0] := 0.00236452;
      W_o[15,1] := 0.63163251;
      W_o[15,2] := 0.04516845;
      W_o[15,3] := -0.19724478;
      W_o[15,4] := -0.66759872;
      W_o[15,5] := 0.38065243;
      W_o[15,6] := 0.64755207;
      W_o[15,7] := 0.26951975;
      W_o[15,8] := -0.49854246;
      W_o[15,9] := -0.37755281;
      W_o[15,10] := 0.25539204;
      W_o[15,11] := -0.14993131;
      W_o[15,12] := 0.57553506;
      W_o[15,13] := -0.03951031;
      W_o[15,14] := 0.02471058;
      W_o[15,15] := -0.23478894;
      W_o[15,16] := 0.31191325;
      W_o[15,17] := 0.02724188;
      W_o[15,18] := 0.33746913;
      W_o[15,19] := -0.03296430;
      W_o[15,20] := -0.88625729;
      W_o[15,21] := 0.50198925;
      W_o[15,22] := -0.01491885;
      W_o[15,23] := 0.39353397;
      W_o[15,24] := 0.29510143;
      W_o[15,25] := 0.44236845;
      W_o[15,26] := -0.03397221;
      W_o[15,27] := -0.45137960;
      W_o[15,28] := 0.26147303;
      W_o[15,29] := -0.10546944;
      W_o[15,30] := 0.30785257;
      W_o[15,31] := -0.10442040;
      W_o[15,32] := 0.27781850;
      W_o[15,33] := -0.00624027;
      W_o[15,34] := 0.29652923;
      W_o[15,35] := -0.21592471;
      W_o[15,36] := 0.05058118;
      W_o[15,37] := 0.00013962;
      W_o[15,38] := 1.00075674;
      W_o[15,39] := 0.55716354;
      R_i[0,0] := -0.11371495;
      R_i[0,1] := -0.00305563;
      R_i[0,2] := 0.44982517;
      R_i[0,3] := 0.40809602;
      R_i[0,4] := 0.49668232;
      R_i[0,5] := 0.26852247;
      R_i[0,6] := 0.58299357;
      R_i[0,7] := 0.30951196;
      R_i[0,8] := 0.58475602;
      R_i[0,9] := 0.44255674;
      R_i[0,10] := 0.16863602;
      R_i[0,11] := -0.31445402;
      R_i[0,12] := 0.01961905;
      R_i[0,13] := 0.39728257;
      R_i[0,14] := 0.35888743;
      R_i[0,15] := 0.12094464;
      R_i[1,0] := -0.03926941;
      R_i[1,1] := -0.22567289;
      R_i[1,2] := -0.18908580;
      R_i[1,3] := -0.40770128;
      R_i[1,4] := 1.58035624;
      R_i[1,5] := -0.53342944;
      R_i[1,6] := -0.07024953;
      R_i[1,7] := 0.42767206;
      R_i[1,8] := -0.66114736;
      R_i[1,9] := 0.46775076;
      R_i[1,10] := -0.07782394;
      R_i[1,11] := -0.44267467;
      R_i[1,12] := 0.19232193;
      R_i[1,13] := 0.63069886;
      R_i[1,14] := -0.44234496;
      R_i[1,15] := -0.14365433;
      R_i[2,0] := -0.10876163;
      R_i[2,1] := -0.00270978;
      R_i[2,2] := 0.21895520;
      R_i[2,3] := -0.58365190;
      R_i[2,4] := -0.07285596;
      R_i[2,5] := 0.04414057;
      R_i[2,6] := 0.29440209;
      R_i[2,7] := -0.56367886;
      R_i[2,8] := 0.02525483;
      R_i[2,9] := 0.21385235;
      R_i[2,10] := 0.14953010;
      R_i[2,11] := 0.47676978;
      R_i[2,12] := 0.35936931;
      R_i[2,13] := -0.47532603;
      R_i[2,14] := -0.06119934;
      R_i[2,15] := -0.18144238;
      R_i[3,0] := -0.34777316;
      R_i[3,1] := -0.02923841;
      R_i[3,2] := -0.01545414;
      R_i[3,3] := 0.67305106;
      R_i[3,4] := 0.52433664;
      R_i[3,5] := 0.12408287;
      R_i[3,6] := 0.36671537;
      R_i[3,7] := 0.40026966;
      R_i[3,8] := 0.66468000;
      R_i[3,9] := 0.16773334;
      R_i[3,10] := 0.19112340;
      R_i[3,11] := -0.51087344;
      R_i[3,12] := 0.11247457;
      R_i[3,13] := -0.26566237;
      R_i[3,14] := 0.38244906;
      R_i[3,15] := -0.15219148;
      R_i[4,0] := 0.00580328;
      R_i[4,1] := 0.66458470;
      R_i[4,2] := -0.75311565;
      R_i[4,3] := 0.00536597;
      R_i[4,4] := -1.54792559;
      R_i[4,5] := -0.47034121;
      R_i[4,6] := -0.23583806;
      R_i[4,7] := 0.20629224;
      R_i[4,8] := 0.50564343;
      R_i[4,9] := 0.17056647;
      R_i[4,10] := -0.12698396;
      R_i[4,11] := -1.01407290;
      R_i[4,12] := 0.52019215;
      R_i[4,13] := -0.14781453;
      R_i[4,14] := -0.18720728;
      R_i[4,15] := -0.01908887;
      R_i[5,0] := -0.57244217;
      R_i[5,1] := 0.07744113;
      R_i[5,2] := 0.07027231;
      R_i[5,3] := 0.15789840;
      R_i[5,4] := 0.23152333;
      R_i[5,5] := 0.13789915;
      R_i[5,6] := -0.36475870;
      R_i[5,7] := -0.19869615;
      R_i[5,8] := -0.04011904;
      R_i[5,9] := -0.05832585;
      R_i[5,10] := -0.04800356;
      R_i[5,11] := -0.20219171;
      R_i[5,12] := -0.02367323;
      R_i[5,13] := 0.18019785;
      R_i[5,14] := 0.07786623;
      R_i[5,15] := -0.41444033;
      R_i[6,0] := -0.48980621;
      R_i[6,1] := -0.08807379;
      R_i[6,2] := 0.72962397;
      R_i[6,3] := 0.53443354;
      R_i[6,4] := -0.33945608;
      R_i[6,5] := 0.02468326;
      R_i[6,6] := -0.59657538;
      R_i[6,7] := -0.15230641;
      R_i[6,8] := -0.06543954;
      R_i[6,9] := 0.06520440;
      R_i[6,10] := -0.09473334;
      R_i[6,11] := 0.06633532;
      R_i[6,12] := 0.55549175;
      R_i[6,13] := -0.56575418;
      R_i[6,14] := 0.12516849;
      R_i[6,15] := -1.21049595;
      R_i[7,0] := 0.09141196;
      R_i[7,1] := -0.29539478;
      R_i[7,2] := -0.04736479;
      R_i[7,3] := 0.63814592;
      R_i[7,4] := -0.17358984;
      R_i[7,5] := 0.02200026;
      R_i[7,6] := -0.54248303;
      R_i[7,7] := 0.41123483;
      R_i[7,8] := 0.08935327;
      R_i[7,9] := 0.21178399;
      R_i[7,10] := 0.37781638;
      R_i[7,11] := -0.24556014;
      R_i[7,12] := -0.25292242;
      R_i[7,13] := 0.36763078;
      R_i[7,14] := -0.16423522;
      R_i[7,15] := 0.30131927;
      R_i[8,0] := -0.43597510;
      R_i[8,1] := 0.53708863;
      R_i[8,2] := -0.01918638;
      R_i[8,3] := 0.06577428;
      R_i[8,4] := -0.23607059;
      R_i[8,5] := 0.04361986;
      R_i[8,6] := 0.43726206;
      R_i[8,7] := 0.31797796;
      R_i[8,8] := -1.00093663;
      R_i[8,9] := -0.33588576;
      R_i[8,10] := 0.94019109;
      R_i[8,11] := -0.48441434;
      R_i[8,12] := -0.02272851;
      R_i[8,13] := 0.18289326;
      R_i[8,14] := -0.01882748;
      R_i[8,15] := -0.06172743;
      R_i[9,0] := -0.51438624;
      R_i[9,1] := 0.06295519;
      R_i[9,2] := 0.30461141;
      R_i[9,3] := 0.03788998;
      R_i[9,4] := 0.13080329;
      R_i[9,5] := -0.35847402;
      R_i[9,6] := 0.69233000;
      R_i[9,7] := -0.27768511;
      R_i[9,8] := 0.00155199;
      R_i[9,9] := -0.09497612;
      R_i[9,10] := 0.19121598;
      R_i[9,11] := -0.42883599;
      R_i[9,12] := 0.09758300;
      R_i[9,13] := 0.28921250;
      R_i[9,14] := 0.13413866;
      R_i[9,15] := -0.65263885;
      R_i[10,0] := -1.24392521;
      R_i[10,1] := 0.68045098;
      R_i[10,2] := 0.94528174;
      R_i[10,3] := -1.11527085;
      R_i[10,4] := -0.62745446;
      R_i[10,5] := -0.47022989;
      R_i[10,6] := 0.90557086;
      R_i[10,7] := 0.78638017;
      R_i[10,8] := 1.25939584;
      R_i[10,9] := 0.48661330;
      R_i[10,10] := -0.23223703;
      R_i[10,11] := -0.88113469;
      R_i[10,12] := -0.14167067;
      R_i[10,13] := 0.25197980;
      R_i[10,14] := 0.71458435;
      R_i[10,15] := -0.03913529;
      R_i[11,0] := -0.29863074;
      R_i[11,1] := 0.74166214;
      R_i[11,2] := -0.54186344;
      R_i[11,3] := -0.02086760;
      R_i[11,4] := 0.44549692;
      R_i[11,5] := -0.15922859;
      R_i[11,6] := 0.25055087;
      R_i[11,7] := -0.38269201;
      R_i[11,8] := 0.16184135;
      R_i[11,9] := 0.41939276;
      R_i[11,10] := 0.02712804;
      R_i[11,11] := -1.18685222;
      R_i[11,12] := 0.20019490;
      R_i[11,13] := 0.15325017;
      R_i[11,14] := -0.32840040;
      R_i[11,15] := -0.28205517;
      R_i[12,0] := -0.28950748;
      R_i[12,1] := 1.09143484;
      R_i[12,2] := -0.05338987;
      R_i[12,3] := 0.29111606;
      R_i[12,4] := 0.16297169;
      R_i[12,5] := -0.16159102;
      R_i[12,6] := 0.51468766;
      R_i[12,7] := 0.03626299;
      R_i[12,8] := 0.08357667;
      R_i[12,9] := 0.27675816;
      R_i[12,10] := -0.27259591;
      R_i[12,11] := -0.94452316;
      R_i[12,12] := 2.16417599;
      R_i[12,13] := -0.04564672;
      R_i[12,14] := -0.94376862;
      R_i[12,15] := -0.37525555;
      R_i[13,0] := -0.37388137;
      R_i[13,1] := -0.43020728;
      R_i[13,2] := 0.06173271;
      R_i[13,3] := -0.32806039;
      R_i[13,4] := -0.27162644;
      R_i[13,5] := 0.35506669;
      R_i[13,6] := -0.05685175;
      R_i[13,7] := 0.51354361;
      R_i[13,8] := 0.16403134;
      R_i[13,9] := -0.26913187;
      R_i[13,10] := -0.38018483;
      R_i[13,11] := 0.12280507;
      R_i[13,12] := 0.54280287;
      R_i[13,13] := 1.70935917;
      R_i[13,14] := 1.01156926;
      R_i[13,15] := -0.42882025;
      R_i[14,0] := 0.23007612;
      R_i[14,1] := -1.01209235;
      R_i[14,2] := 0.63614035;
      R_i[14,3] := 0.05786986;
      R_i[14,4] := -0.45537889;
      R_i[14,5] := -0.66792619;
      R_i[14,6] := -0.40340808;
      R_i[14,7] := 0.00973069;
      R_i[14,8] := 1.01184237;
      R_i[14,9] := -0.35905090;
      R_i[14,10] := 0.33358613;
      R_i[14,11] := -0.82171744;
      R_i[14,12] := -0.64750588;
      R_i[14,13] := -0.20203376;
      R_i[14,14] := 3.03613806;
      R_i[14,15] := -0.17449842;
      R_i[15,0] := -0.04125203;
      R_i[15,1] := 0.67002559;
      R_i[15,2] := 1.07735050;
      R_i[15,3] := 0.28749722;
      R_i[15,4] := -0.03804383;
      R_i[15,5] := 0.07771160;
      R_i[15,6] := 0.64223152;
      R_i[15,7] := 0.28548393;
      R_i[15,8] := 0.24192756;
      R_i[15,9] := 0.00585660;
      R_i[15,10] := 0.62889910;
      R_i[15,11] := -0.83460343;
      R_i[15,12] := 0.24951389;
      R_i[15,13] := -0.46169642;
      R_i[15,14] := 0.85477173;
      R_i[15,15] := -1.05970228;
      R_f[0,0] := 0.32337135;
      R_f[0,1] := -0.64154255;
      R_f[0,2] := 0.44366962;
      R_f[0,3] := -0.16911837;
      R_f[0,4] := -0.22606935;
      R_f[0,5] := 0.40707147;
      R_f[0,6] := 0.99587154;
      R_f[0,7] := -0.61522830;
      R_f[0,8] := -0.16690622;
      R_f[0,9] := 0.11400585;
      R_f[0,10] := -1.30126393;
      R_f[0,11] := 0.68435878;
      R_f[0,12] := 0.25505054;
      R_f[0,13] := -0.50005764;
      R_f[0,14] := 1.89920795;
      R_f[0,15] := 0.31197056;
      R_f[1,0] := -0.10116166;
      R_f[1,1] := 3.47733283;
      R_f[1,2] := -0.23958448;
      R_f[1,3] := 0.25761580;
      R_f[1,4] := 0.64858228;
      R_f[1,5] := 0.25520656;
      R_f[1,6] := 0.47342876;
      R_f[1,7] := 0.44394684;
      R_f[1,8] := 0.08832169;
      R_f[1,9] := -0.07672439;
      R_f[1,10] := -0.11365046;
      R_f[1,11] := -0.12767753;
      R_f[1,12] := 0.15301596;
      R_f[1,13] := 0.10815746;
      R_f[1,14] := -0.00451868;
      R_f[1,15] := 0.16956279;
      R_f[2,0] := 0.88069433;
      R_f[2,1] := -0.43075773;
      R_f[2,2] := -0.28541803;
      R_f[2,3] := 0.77957338;
      R_f[2,4] := 0.49963999;
      R_f[2,5] := 0.15426520;
      R_f[2,6] := 0.22863509;
      R_f[2,7] := -0.74026376;
      R_f[2,8] := -0.68504810;
      R_f[2,9] := -0.34440613;
      R_f[2,10] := -0.51462018;
      R_f[2,11] := 0.52031350;
      R_f[2,12] := -0.29210886;
      R_f[2,13] := -0.75812620;
      R_f[2,14] := 0.24005084;
      R_f[2,15] := 0.06470054;
      R_f[3,0] := -1.01638353;
      R_f[3,1] := -0.01572494;
      R_f[3,2] := 1.12268722;
      R_f[3,3] := -1.07652342;
      R_f[3,4] := -0.22190276;
      R_f[3,5] := 0.38419157;
      R_f[3,6] := 0.65128225;
      R_f[3,7] := 1.68439031;
      R_f[3,8] := 0.77879173;
      R_f[3,9] := -0.13034230;
      R_f[3,10] := 0.10257917;
      R_f[3,11] := 0.06301130;
      R_f[3,12] := -0.26139963;
      R_f[3,13] := 0.08574831;
      R_f[3,14] := 0.58179146;
      R_f[3,15] := -0.16947731;
      R_f[4,0] := -0.09817147;
      R_f[4,1] := -0.86730129;
      R_f[4,2] := 0.11236032;
      R_f[4,3] := -0.05304767;
      R_f[4,4] := -0.16176023;
      R_f[4,5] := -0.43156531;
      R_f[4,6] := -0.15450424;
      R_f[4,7] := -0.04651795;
      R_f[4,8] := -0.77932215;
      R_f[4,9] := 0.20782343;
      R_f[4,10] := 0.16769727;
      R_f[4,11] := 0.33256632;
      R_f[4,12] := 0.15797095;
      R_f[4,13] := 0.73622912;
      R_f[4,14] := 0.01762660;
      R_f[4,15] := -0.67344528;
      R_f[5,0] := 1.16960347;
      R_f[5,1] := -0.73157996;
      R_f[5,2] := 0.41226324;
      R_f[5,3] := 0.02196453;
      R_f[5,4] := 0.35487083;
      R_f[5,5] := 0.18895856;
      R_f[5,6] := 0.30451256;
      R_f[5,7] := 0.92117321;
      R_f[5,8] := -0.48577240;
      R_f[5,9] := -0.98202080;
      R_f[5,10] := -0.51303148;
      R_f[5,11] := 0.26235431;
      R_f[5,12] := -0.22034658;
      R_f[5,13] := -1.83764625;
      R_f[5,14] := -0.65874094;
      R_f[5,15] := -0.29308036;
      R_f[6,0] := -0.39891392;
      R_f[6,1] := -0.75305557;
      R_f[6,2] := 1.69584787;
      R_f[6,3] := -0.16370860;
      R_f[6,4] := 0.25405717;
      R_f[6,5] := 0.02853256;
      R_f[6,6] := 0.15147270;
      R_f[6,7] := -1.13414180;
      R_f[6,8] := -0.99144781;
      R_f[6,9] := -0.44909641;
      R_f[6,10] := -0.64757788;
      R_f[6,11] := -0.02062916;
      R_f[6,12] := 0.33514625;
      R_f[6,13] := 0.30901858;
      R_f[6,14] := 0.61397654;
      R_f[6,15] := 0.76879233;
      R_f[7,0] := -0.27052191;
      R_f[7,1] := 0.04162847;
      R_f[7,2] := 3.14724135;
      R_f[7,3] := -0.33119497;
      R_f[7,4] := -0.58844078;
      R_f[7,5] := -0.36365259;
      R_f[7,6] := -0.91634971;
      R_f[7,7] := 0.35394892;
      R_f[7,8] := 0.28250608;
      R_f[7,9] := 0.49327499;
      R_f[7,10] := 1.35347533;
      R_f[7,11] := -1.12448680;
      R_f[7,12] := -0.59189665;
      R_f[7,13] := 1.29001379;
      R_f[7,14] := -0.55096096;
      R_f[7,15] := 0.86654115;
      R_f[8,0] := 0.36559653;
      R_f[8,1] := -1.38739824;
      R_f[8,2] := 0.64030659;
      R_f[8,3] := 0.45218420;
      R_f[8,4] := 0.42656797;
      R_f[8,5] := -0.34682584;
      R_f[8,6] := -1.10001183;
      R_f[8,7] := -0.66935474;
      R_f[8,8] := -3.06901670;
      R_f[8,9] := 0.16576712;
      R_f[8,10] := 0.78494203;
      R_f[8,11] := -0.43459168;
      R_f[8,12] := -1.43488169;
      R_f[8,13] := 0.13381413;
      R_f[8,14] := -0.79348296;
      R_f[8,15] := -0.22492136;
      R_f[9,0] := -0.15259695;
      R_f[9,1] := -1.49991405;
      R_f[9,2] := 1.10876131;
      R_f[9,3] := -0.52977806;
      R_f[9,4] := -0.68868691;
      R_f[9,5] := -1.67290866;
      R_f[9,6] := 2.63343525;
      R_f[9,7] := -1.82854438;
      R_f[9,8] := -0.74066204;
      R_f[9,9] := 1.52620482;
      R_f[9,10] := 0.47460184;
      R_f[9,11] := 1.38148880;
      R_f[9,12] := -0.60541850;
      R_f[9,13] := 0.79266793;
      R_f[9,14] := 0.32717809;
      R_f[9,15] := -1.00011170;
      R_f[10,0] := 2.16440725;
      R_f[10,1] := -0.69953722;
      R_f[10,2] := 0.66533321;
      R_f[10,3] := 1.18175888;
      R_f[10,4] := -0.29653463;
      R_f[10,5] := -0.10375768;
      R_f[10,6] := 0.02757812;
      R_f[10,7] := -0.96818727;
      R_f[10,8] := -0.46075854;
      R_f[10,9] := -0.54467458;
      R_f[10,10] := 0.78059703;
      R_f[10,11] := -0.76885021;
      R_f[10,12] := -1.05606675;
      R_f[10,13] := -0.19888546;
      R_f[10,14] := 0.01456859;
      R_f[10,15] := 0.37021348;
      R_f[11,0] := 0.24349366;
      R_f[11,1] := -0.17989418;
      R_f[11,2] := 0.23558758;
      R_f[11,3] := -0.66829973;
      R_f[11,4] := -0.50071466;
      R_f[11,5] := -0.57912046;
      R_f[11,6] := 0.12530079;
      R_f[11,7] := -0.76207477;
      R_f[11,8] := -0.57875133;
      R_f[11,9] := 0.02648440;
      R_f[11,10] := 0.43179271;
      R_f[11,11] := -1.22257721;
      R_f[11,12] := -0.03755289;
      R_f[11,13] := -0.12284968;
      R_f[11,14] := 0.06467830;
      R_f[11,15] := 0.26499867;
      R_f[12,0] := -0.02412502;
      R_f[12,1] := -0.41788927;
      R_f[12,2] := 0.22505651;
      R_f[12,3] := 0.24685313;
      R_f[12,4] := -0.26033589;
      R_f[12,5] := 0.55886257;
      R_f[12,6] := 0.35019273;
      R_f[12,7] := 0.06464690;
      R_f[12,8] := 0.38953316;
      R_f[12,9] := 0.40905604;
      R_f[12,10] := 0.16141498;
      R_f[12,11] := -0.05112006;
      R_f[12,12] := 1.49376774;
      R_f[12,13] := 0.31314605;
      R_f[12,14] := 0.45734319;
      R_f[12,15] := 0.38003021;
      R_f[13,0] := 0.59145856;
      R_f[13,1] := -0.35116604;
      R_f[13,2] := 0.82912683;
      R_f[13,3] := 0.20134470;
      R_f[13,4] := 0.82876003;
      R_f[13,5] := 0.89772320;
      R_f[13,6] := 1.65778053;
      R_f[13,7] := 0.49528536;
      R_f[13,8] := -0.85102677;
      R_f[13,9] := -0.78163058;
      R_f[13,10] := 0.37120518;
      R_f[13,11] := 0.77949518;
      R_f[13,12] := -0.15100223;
      R_f[13,13] := -0.17492811;
      R_f[13,14] := -0.00674355;
      R_f[13,15] := -0.65944511;
      R_f[14,0] := -0.03948923;
      R_f[14,1] := -0.36825284;
      R_f[14,2] := 1.24439776;
      R_f[14,3] := -0.53740013;
      R_f[14,4] := -0.42868876;
      R_f[14,5] := 0.26089478;
      R_f[14,6] := 0.48867851;
      R_f[14,7] := 1.19528174;
      R_f[14,8] := 0.15456729;
      R_f[14,9] := -1.14040160;
      R_f[14,10] := 0.05182516;
      R_f[14,11] := -0.21726616;
      R_f[14,12] := 0.17021520;
      R_f[14,13] := -0.64748013;
      R_f[14,14] := 1.38772130;
      R_f[14,15] := 0.23228650;
      R_f[15,0] := 0.31530645;
      R_f[15,1] := -0.98082370;
      R_f[15,2] := 0.22649910;
      R_f[15,3] := -0.29767367;
      R_f[15,4] := 0.54684836;
      R_f[15,5] := 0.77809179;
      R_f[15,6] := 2.00395179;
      R_f[15,7] := 2.35574341;
      R_f[15,8] := -0.17023613;
      R_f[15,9] := -0.38121098;
      R_f[15,10] := 1.06925368;
      R_f[15,11] := -0.30545777;
      R_f[15,12] := -0.43472868;
      R_f[15,13] := -1.11482680;
      R_f[15,14] := 0.32454339;
      R_f[15,15] := -1.33770871;
      R_g[0,0] := -2.80543303;
      R_g[0,1] := 0.09675837;
      R_g[0,2] := 0.04763355;
      R_g[0,3] := 0.16134985;
      R_g[0,4] := -0.04916951;
      R_g[0,5] := 0.06786807;
      R_g[0,6] := 0.07195669;
      R_g[0,7] := 0.18796267;
      R_g[0,8] := 0.02096096;
      R_g[0,9] := -0.05091592;
      R_g[0,10] := 0.17113523;
      R_g[0,11] := 0.09710391;
      R_g[0,12] := -0.19285078;
      R_g[0,13] := 0.04608029;
      R_g[0,14] := 0.37757719;
      R_g[0,15] := -0.05004899;
      R_g[1,0] := 0.08712953;
      R_g[1,1] := -1.28173816;
      R_g[1,2] := 0.48629102;
      R_g[1,3] := -0.10185467;
      R_g[1,4] := 0.59114659;
      R_g[1,5] := 0.38262466;
      R_g[1,6] := 0.04029783;
      R_g[1,7] := 0.06582787;
      R_g[1,8] := -0.06752597;
      R_g[1,9] := -0.22948581;
      R_g[1,10] := -0.12531509;
      R_g[1,11] := -0.20673551;
      R_g[1,12] := -0.05208173;
      R_g[1,13] := 0.18107648;
      R_g[1,14] := 0.05905702;
      R_g[1,15] := -0.06634986;
      R_g[2,0] := -0.25491390;
      R_g[2,1] := -0.05303259;
      R_g[2,2] := -3.25826526;
      R_g[2,3] := 0.22390363;
      R_g[2,4] := 0.08010214;
      R_g[2,5] := 0.12519346;
      R_g[2,6] := -0.12813619;
      R_g[2,7] := 0.03709217;
      R_g[2,8] := -0.05339420;
      R_g[2,9] := -0.18383153;
      R_g[2,10] := 0.01583981;
      R_g[2,11] := 0.12061389;
      R_g[2,12] := 0.02361463;
      R_g[2,13] := 0.11624731;
      R_g[2,14] := 0.16856082;
      R_g[2,15] := -0.04670952;
      R_g[3,0] := -0.34998056;
      R_g[3,1] := 0.71455550;
      R_g[3,2] := -0.79799318;
      R_g[3,3] := -2.84151006;
      R_g[3,4] := 0.15804654;
      R_g[3,5] := -0.08033045;
      R_g[3,6] := -0.14524731;
      R_g[3,7] := 0.22259524;
      R_g[3,8] := 0.07427457;
      R_g[3,9] := 0.37250251;
      R_g[3,10] := -0.30889195;
      R_g[3,11] := -0.23224294;
      R_g[3,12] := 0.67339027;
      R_g[3,13] := 0.18020143;
      R_g[3,14] := -0.04057474;
      R_g[3,15] := -0.17805941;
      R_g[4,0] := 0.45585641;
      R_g[4,1] := 0.26910168;
      R_g[4,2] := 0.24799341;
      R_g[4,3] := 0.18304951;
      R_g[4,4] := -2.64359164;
      R_g[4,5] := -0.18548726;
      R_g[4,6] := 0.57962537;
      R_g[4,7] := -0.23603684;
      R_g[4,8] := 0.39961720;
      R_g[4,9] := -0.08552616;
      R_g[4,10] := -0.35479608;
      R_g[4,11] := 0.02176627;
      R_g[4,12] := -0.16954437;
